RoboDK station: RobotPrint_Printhead_cbeam 1.rdk

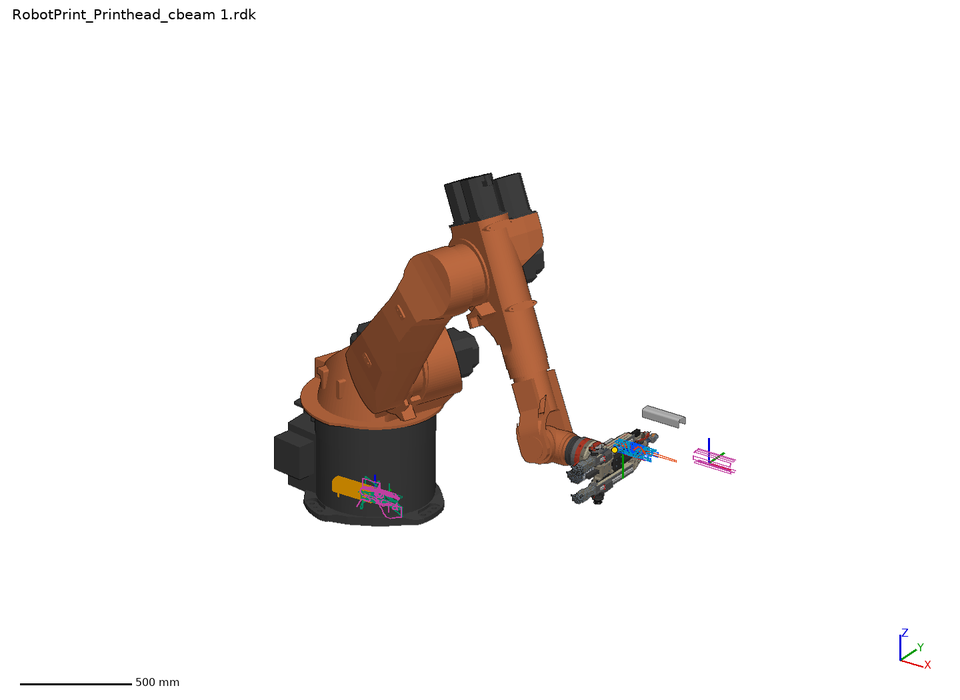
[picture v0: the station drawn from its stored meshes, robots at their saved joint values, targets as dots, program paths as lines]
Station RobotPrinter_Printhead (saved by RoboDK 5.8.0). Poses are relative to the parent item; angles as X-Y-Z fixed-axis rotations.
  - frame KUKA KR 30 HA Base at (0, 0, 0) mm
    - robot KUKA KR 30 HA: 6 axes, payload 30 kg, reach 2033 mm, repeatability 0.05 mm, weight 665 kg
        modified DH rows (alpha deg, a mm, theta deg, d mm): 0, 0, 0, 815; -90, 350, 0, 0; 0, 850, -90, 0; -90, 145, 0, 820; 90, 0, 0, 0; -90, 0, 180, 170
        joint limits [-185, -135, -120, -350, -119, -350] to [185, 35, 158, 350, 119, 350]; home [0, -90, 90, 0, 0, 0]; saved at [20.826, -52.741, 114.474, 203.359, 63.728, -280.823]
      - tool PlasticPos800, TCP at (350.64, -42.92, 173.8) mm
      - tool PlasticPos1200, TCP at (391.44, -42.9, 173.32) mm
      - tool FiberPos800, TCP at (355.38, 32.86, 175) mm, rotated rx 0 ry 90 rz 0 deg
      - tool FiberPos1200, TCP at (394.69, 33.62, 175.94) mm
      - tool Printheady, TCP at (0, 0, 200) mm, size 292.2 x 550.3 x 343.3 mm, geometry from CAD_Printheady.step
      - tool TOOL 0, TCP at (0, 0, 0) mm
    - frame PrintbedOrigin at (1792.66, 35.63, 669.38) mm
    - frame Reference SW at (1415.36, -92.38, 659.99) mm, rotated rx -90 ry 0 rz 0 deg
      - object C-Beam-5mm-200mm RoboDK-Test at (300, -210, 0) mm, size 200 x 40 x 50 mm, geometry from C-Beam-5mm-200mm RoboDK-Test.stl
      - object C-Beam-5mm-200mm RoboDK-Test 1 at (0, 0, 0) mm, size 200 x 50 x 50 mm, geometry from C-Beam-5mm-200mm RoboDK-Test 1.stl
      - object CBL1-2 at (0, 0, 0) mm
      - object CBL2-2 at (0, 0, 0) mm
      - object CBL1 at (0, 0, 0) mm
    - frame BASE 0 at (0, 0, 0) mm
  - machining project CBL1-2 Settings: rotZ(0) | rotX(0)*rotY(0) | onStart | onPathStart | onApproach | onPoint | onRetract | onFinish | SetRPM(%1) | SetTool(%1) | Extruder(%1) | default | default | OutOnMov(%1) | OutOffMov(%1) | onPathFinish | M_RunCode(%1)
  - program CBL1-2 (86 instructions, listed below)
  - machining project CBL2-2 Settings: rotZ(0) | rotX(0)*rotY(0) | rotz(0) | onStart | onPathStart | onApproach | onPoint | onRetract | onFinish | SetRPM(%1) | SetTool(%1) | Extruder(%1) | default | default | OutOnMov(%1) | OutOffMov(%1) | onPathFinish | M_RunCode(%1)
  - program CBL2-2 (24 instructions, listed below)
  - program CBL12 (41 instructions, listed below)
  - program CBL12 (44 instructions, listed below)
  - program CBL12 (39 instructions, listed below)
  - machining project Pfad3 Einstellungen: rotZ(0) | rotX(0)*rotY(0) | onStart | onPathStart | onApproach | onPoint | onRetract | onFinish | SetRPM(%1) | SetTool(%1) | Extruder(%1) | default | default | OutOnMov(%1) | OutOffMov(%1) | onPathFinish | M_RunCode(%1)
  - program Pfad3 (95 instructions, listed below)
  - program TP12Layers (5237 instructions, listed below)
  - machining project CBL1 Settings: rotZ(0) | rotX(0)*rotY(0) | onStart | onPathStart | onApproach | onPoint | onRetract | onFinish | SetRPM(%1) | SetTool(%1) | Extruder(%1) | default | default | OutOnMov(%1) | OutOffMov(%1) | onPathFinish | M_RunCode(%1)
  - program CBL1 (341 instructions, listed below)
  - machining project Pfad5 Einstellungen: rotZ(0) | rotX(0)*rotY(0) | onStart | onPathStart | onApproach | onPoint | onRetract | onFinish | SetRPM(%1) | SetTool(%1) | Extruder(%1) | default | default | OutOnMov(%1) | OutOffMov(%1) | onPathFinish | M_RunCode(%1)
  - program Pfad5 (148 instructions, listed below)
  - machining project Pfad6 Einstellungen: rotZ(0) | rotX(0)*rotY(0) | onStart | onPathStart | onApproach | onPoint | onRetract | onFinish | SetRPM(%1) | SetTool(%1) | Extruder(%1) | default | default | OutOnMov(%1) | OutOffMov(%1) | onPathFinish | M_RunCode(%1)
  - program Pfad6 (33 instructions, listed below)
  - program CFSteer (1006 instructions, listed below)
  - program CFLines (937 instructions, listed below)
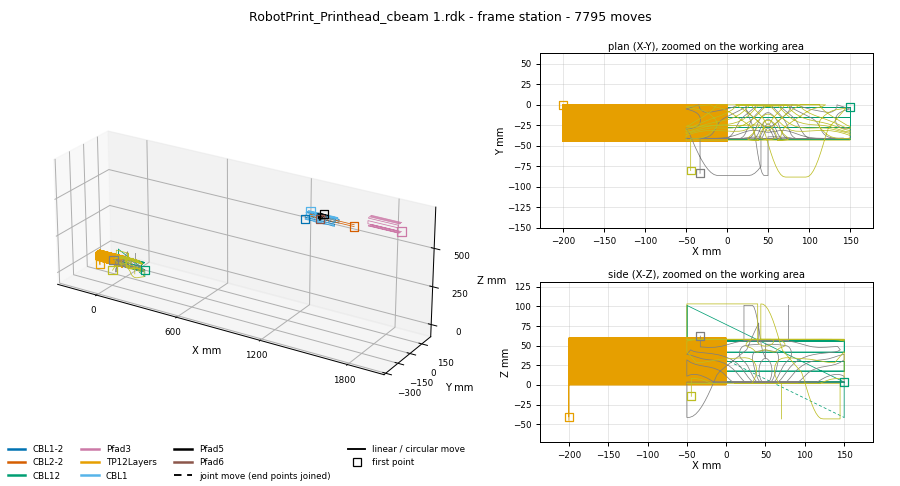
[picture p0: tool path of RobotPrint_Printhead_cbeam 1.rdk in frame station, 7795 of 7795 moves have a stored position in this frame; points joined in program order, loops and branches not executed]

--- program CBL1-2 (robot KUKA KR 30 HA) ---
  Glatt(1)
  Sollgeschwindigkeit (1000.0 mm/s)
  Referenz erstellen.: Reference SW
  Werkzeug setzen: FiberPos800
  Anzeigen FiberPos800
  MoveJ 1 to (-50, -3, 3.75) mm, rotated rx 180 ry 0 rz -90 deg; joints [-10.801, -58.742, 109.357, 0, 39.385, 79.199]
  MoveL 2 to (-50, -3, 3.75) mm, rotated rx 180 ry 0 rz -90 deg; joints [-10.801, -58.742, 109.357, 0, 39.385, 79.199]
  MoveL 3 to (-50, -3, 3.75) mm, rotated rx 180 ry 0 rz -90 deg; joints [-10.801, -58.742, 109.357, 0, 39.385, 79.199]
  MoveL 4 to (-50, -3, 3.75) mm, rotated rx 180 ry 0 rz -90 deg; joints [-10.801, -58.742, 109.357, 0, 39.385, 79.199]
  Sollgeschwindigkeit (50.0 mm/s)
  MoveL 5 to (150, -3, 3.75) mm, rotated rx -180 ry 0 rz -90 deg; joints [-9.475, -48.064, 90.596, 0, 47.468, 80.525]
  Sollgeschwindigkeit (1000.0 mm/s)
  MoveL 6 to (150, -3, 3.75) mm, rotated rx -180 ry 0 rz -90 deg; joints [-9.475, -48.064, 90.596, 0, 47.468, 80.525]
  MoveL 7 to (150, -3, 3.75) mm, rotated rx -180 ry 0 rz -90 deg; joints [-9.475, -48.064, 90.596, 0, 47.468, 80.525]
  Sollgeschwindigkeit (1000.0 mm/s)
  MoveL 8 to (150, -15, 3.75) mm, rotated rx -180 ry 0 rz -90 deg; joints [-9.475, -48.501, 90.408, 0, 48.093, 80.525]
  MoveL 9 to (150, -15, 3.75) mm, rotated rx -180 ry 0 rz -90 deg; joints [-9.475, -48.501, 90.408, 0, 48.093, 80.525]
  MoveL 10 to (150, -15, 3.75) mm, rotated rx -180 ry 0 rz -90 deg; joints [-9.475, -48.501, 90.408, 0, 48.093, 80.525]
  Sollgeschwindigkeit (50.0 mm/s)
  MoveL 11 to (-50, -15, 3.75) mm, rotated rx 180 ry 0 rz -90 deg; joints [-10.801, -59.271, 109.17, 0, 40.102, 79.199]
  Sollgeschwindigkeit (1000.0 mm/s)
  MoveL 12 to (-50, -15, 3.75) mm, rotated rx 180 ry 0 rz -90 deg; joints [-10.801, -59.271, 109.17, 0, 40.102, 79.199]
  MoveL 13 to (-50, -15, 3.75) mm, rotated rx 180 ry 0 rz -90 deg; joints [-10.801, -59.271, 109.17, 0, 40.102, 79.199]
  Sollgeschwindigkeit (1000.0 mm/s)
  MoveL 14 to (-50, -27, 3.75) mm, rotated rx 180 ry 0 rz -90 deg; joints [-10.801, -59.792, 108.97, 0, 40.822, 79.199]
  MoveL 15 to (-50, -27, 3.75) mm, rotated rx 180 ry 0 rz -90 deg; joints [-10.801, -59.792, 108.97, 0, 40.822, 79.199]
  MoveL 16 to (-50, -27, 3.75) mm, rotated rx 180 ry 0 rz -90 deg; joints [-10.801, -59.792, 108.97, 0, 40.822, 79.199]
  Sollgeschwindigkeit (50.0 mm/s)
  MoveL 17 to (150, -27, 3.75) mm, rotated rx -180 ry 0 rz -90 deg; joints [-9.475, -48.931, 90.208, 0, 48.722, 80.525]
  Sollgeschwindigkeit (1000.0 mm/s)
  MoveL 18 to (150, -27, 3.75) mm, rotated rx -180 ry 0 rz -90 deg; joints [-9.475, -48.931, 90.208, 0, 48.722, 80.525]
  MoveL 19 to (150, -27, 3.75) mm, rotated rx -180 ry 0 rz -90 deg; joints [-9.475, -48.931, 90.208, 0, 48.722, 80.525]
  Sollgeschwindigkeit (1000.0 mm/s)
  MoveL 20 to (150, -41.25, 18) mm, rotated rx -180 ry 0 rz -90 deg; joints [-9.972, -49.289, 89.704, 0, 49.585, 80.028]
  MoveL 21 to (150, -41.25, 18) mm, rotated rx -180 ry 0 rz -90 deg; joints [-9.972, -49.289, 89.704, 0, 49.585, 80.028]
  MoveL 22 to (150, -41.25, 18) mm, rotated rx -180 ry 0 rz -90 deg; joints [-9.972, -49.289, 89.704, 0, 49.585, 80.028]
  Sollgeschwindigkeit (50.0 mm/s)
  MoveL 23 to (-50, -41.25, 18) mm, rotated rx -180 ry 0 rz -90 deg; joints [-11.363, -60.254, 108.477, 0, 41.777, 78.637]
  Sollgeschwindigkeit (1000.0 mm/s)
  MoveL 24 to (-50, -41.25, 18) mm, rotated rx -180 ry 0 rz -90 deg; joints [-11.363, -60.254, 108.477, 0, 41.777, 78.637]
  MoveL 25 to (-50, -41.25, 18) mm, rotated rx -180 ry 0 rz -90 deg; joints [-11.363, -60.254, 108.477, 0, 41.777, 78.637]
  Sollgeschwindigkeit (1000.0 mm/s)
  MoveL 26 to (-50, -41.25, 30) mm, rotated rx 180 ry 0 rz -90 deg; joints [-11.835, -60.125, 108.264, 0, 41.86, 78.165]
  MoveL 27 to (-50, -41.25, 30) mm, rotated rx 180 ry 0 rz -90 deg; joints [-11.835, -60.125, 108.264, 0, 41.86, 78.165]
  MoveL 28 to (-50, -41.25, 30) mm, rotated rx 180 ry 0 rz -90 deg; joints [-11.835, -60.125, 108.264, 0, 41.86, 78.165]
  Sollgeschwindigkeit (50.0 mm/s)
  MoveL 29 to (150, -41.25, 30) mm, rotated rx -180 ry 0 rz -90 deg; joints [-10.388, -49.164, 89.482, 0, 49.682, 79.612]
  Sollgeschwindigkeit (1000.0 mm/s)
  MoveL 30 to (150, -41.25, 30) mm, rotated rx -180 ry 0 rz -90 deg; joints [-10.388, -49.164, 89.482, 0, 49.682, 79.612]
  MoveL 31 to (150, -41.25, 30) mm, rotated rx -180 ry 0 rz -90 deg; joints [-10.388, -49.164, 89.482, 0, 49.682, 79.612]
  Sollgeschwindigkeit (1000.0 mm/s)
  MoveL 32 to (150, -41.25, 42) mm, rotated rx 180 ry 0 rz -90 deg; joints [-10.804, -49.033, 89.25, 0, 49.783, 79.196]
  MoveL 33 to (150, -41.25, 42) mm, rotated rx 180 ry 0 rz -90 deg; joints [-10.804, -49.033, 89.25, 0, 49.783, 79.196]
  MoveL 34 to (150, -41.25, 42) mm, rotated rx 180 ry 0 rz -90 deg; joints [-10.804, -49.033, 89.25, 0, 49.783, 79.196]
  Sollgeschwindigkeit (50.0 mm/s)
  MoveL 35 to (-50, -41.25, 42) mm, rotated rx -180 ry 0 rz -90 deg; joints [-12.305, -59.99, 108.043, 0, 41.947, 77.695]
  Sollgeschwindigkeit (1000.0 mm/s)
  MoveL 36 to (-50, -41.25, 42) mm, rotated rx -180 ry 0 rz -90 deg; joints [-12.305, -59.99, 108.043, 0, 41.947, 77.695]
  MoveL 37 to (-50, -41.25, 42) mm, rotated rx -180 ry 0 rz -90 deg; joints [-12.305, -59.99, 108.043, 0, 41.947, 77.695]
  Sollgeschwindigkeit (1000.0 mm/s)
  MoveL 38 to (-50, -27, 56.25) mm, rotated rx 180 ry 0 rz -90 deg; joints [-12.862, -59.222, 108.019, 0, 41.202, 77.138]
  MoveL 39 to (-50, -27, 56.25) mm, rotated rx 180 ry 0 rz -90 deg; joints [-12.862, -59.222, 108.019, 0, 41.202, 77.138]
  MoveL 40 to (-50, -27, 56.25) mm, rotated rx 180 ry 0 rz -90 deg; joints [-12.862, -59.222, 108.019, 0, 41.202, 77.138]
  Sollgeschwindigkeit (50.0 mm/s)
  MoveL 41 to (150, -27, 56.25) mm, rotated rx -180 ry 0 rz -90 deg; joints [-11.296, -48.375, 89.215, 0, 49.16, 78.704]
  Sollgeschwindigkeit (1000.0 mm/s)
  MoveL 42 to (150, -27, 56.25) mm, rotated rx -180 ry 0 rz -90 deg; joints [-11.296, -48.375, 89.215, 0, 49.16, 78.704]
  MoveL 43 to (150, -27, 56.25) mm, rotated rx -180 ry 0 rz -90 deg; joints [-11.296, -48.375, 89.215, 0, 49.16, 78.704]
  Sollgeschwindigkeit (1000.0 mm/s)
  MoveL 44 to (150, -15, 56.25) mm, rotated rx -180 ry 0 rz -90 deg; joints [-11.296, -47.95, 89.416, 0, 48.534, 78.704]
  MoveL 45 to (150, -15, 56.25) mm, rotated rx -180 ry 0 rz -90 deg; joints [-11.296, -47.95, 89.416, 0, 48.534, 78.704]
  MoveL 46 to (150, -15, 56.25) mm, rotated rx -180 ry 0 rz -90 deg; joints [-11.296, -47.95, 89.416, 0, 48.534, 78.704]
  Sollgeschwindigkeit (50.0 mm/s)
  MoveL 47 to (-50, -15, 56.25) mm, rotated rx 180 ry 0 rz -90 deg; joints [-12.862, -58.706, 108.219, 0, 40.488, 77.138]
  Sollgeschwindigkeit (1000.0 mm/s)
  MoveL 48 to (-50, -15, 56.25) mm, rotated rx 180 ry 0 rz -90 deg; joints [-12.862, -58.706, 108.219, 0, 40.488, 77.138]
  MoveL 49 to (-50, -15, 56.25) mm, rotated rx 180 ry 0 rz -90 deg; joints [-12.862, -58.706, 108.219, 0, 40.488, 77.138]
  Sollgeschwindigkeit (1000.0 mm/s)
  MoveL 50 to (-50, -3, 56.25) mm, rotated rx 180 ry 0 rz -90 deg; joints [-12.862, -58.183, 108.406, 0, 39.777, 77.138]
  MoveL 51 to (-50, -3, 56.25) mm, rotated rx 180 ry 0 rz -90 deg; joints [-12.862, -58.183, 108.406, 0, 39.777, 77.138]
  MoveL 52 to (-50, -3, 56.25) mm, rotated rx 180 ry 0 rz -90 deg; joints [-12.862, -58.183, 108.406, 0, 39.777, 77.138]
  Sollgeschwindigkeit (50.0 mm/s)
  MoveL 53 to (150, -3, 56.25) mm, rotated rx -180 ry 0 rz -90 deg; joints [-11.296, -47.517, 89.605, 0, 47.912, 78.704]
  Sollgeschwindigkeit (1000.0 mm/s)
  MoveL 54 to (150, -3, 56.25) mm, rotated rx -180 ry 0 rz -90 deg; joints [-11.296, -47.517, 89.605, 0, 47.912, 78.704]
  MoveL 55 to (150, -3, 56.25) mm, rotated rx -180 ry 0 rz -90 deg; joints [-11.296, -47.517, 89.605, 0, 47.912, 78.704]

--- program CBL2-2 (robot KUKA KR 30 HA) ---
  Glatt(1)
  Sollgeschwindigkeit (1000.0 mm/s)
  Referenz erstellen.: Reference SW
  Werkzeug setzen: FiberPos800
  Anzeigen FiberPos800
  MoveJ 1 to (250, -3, 58.75) mm, rotated rx 90 ry 0 rz -90 deg; joints [1.885, -7.943, 13.331, 0, 84.613, 1.885]
  MoveL 2 to (250, -3, 58.75) mm, rotated rx 90 ry 0 rz -90 deg; joints [1.885, -7.943, 13.331, 0, 84.613, 1.885]
  MoveL 3 to (150, -3, 58.75) mm, rotated rx 90 ry 0 rz -90 deg; joints [1.983, -26.347, 49.734, 0, 66.613, 1.983]
  MoveL 4 to (150, -3, 58.75) mm, rotated rx 90 ry 0 rz -90 deg; joints [1.983, -26.347, 49.734, 0, 66.613, 1.983]
  Sollgeschwindigkeit (50.0 mm/s)
  MoveL 5 to (-50, -3, 58.75) mm, rotated rx 90 ry 0 rz -90 deg; joints [2.213, -41.91, 79.315, 0, 52.595, 2.213]
  Sollgeschwindigkeit (1000.0 mm/s)
  MoveL 6 to (-50, -3, 58.75) mm, rotated rx 90 ry 0 rz -90 deg; joints [2.213, -41.91, 79.315, 0, 52.595, 2.213]
  MoveL 7 to (50, -3, 58.75) mm, rotated rx 90 ry 0 rz -90 deg; joints [2.091, -35.006, 66.355, 0, 58.651, 2.091]
  Sollgeschwindigkeit (1000.0 mm/s)
  MoveL 8 to (50, -15, 58.75) mm, rotated rx 90 ry 0 rz -90 deg; joints [2.091, -35.355, 66.132, 0, 59.223, 2.091]
  MoveL 9 to (-50, -15, 58.75) mm, rotated rx 90 ry 0 rz -90 deg; joints [2.213, -42.303, 79.116, 0, 53.187, 2.213]
  MoveL 10 to (-50, -15, 58.75) mm, rotated rx 90 ry 0 rz -90 deg; joints [2.213, -42.303, 79.116, 0, 53.187, 2.213]
  Sollgeschwindigkeit (50.0 mm/s)
  MoveL 11 to (150, -15, 58.75) mm, rotated rx 90 ry 0 rz -90 deg; joints [1.983, -26.634, 49.443, 0, 67.192, 1.983]
  Sollgeschwindigkeit (1000.0 mm/s)
  MoveL 12 to (150, -15, 58.75) mm, rotated rx 90 ry 0 rz -90 deg; joints [1.983, -26.634, 49.443, 0, 67.192, 1.983]
  MoveL 13 to (250, -15, 58.75) mm, rotated rx 90 ry -20 rz -90 deg; joints [-1.516, -8.156, 13.591, 20.06, 85.412, -3.287]
  Sollgeschwindigkeit (1000.0 mm/s)

--- program CBL12 (robot KUKA KR 30 HA) ---
  BAS (#INITMOV,0)
  BAS (#VEL_PTP,100)
  BAS (#ACC_PTP,20)
  Sollgeschwindigkeit (200.0 mm/s)
  Werkzeug setzen: TOOL 0
  Referenz erstellen.: BASE 0
  $ADVANCE = 5
  $APO.CPTP = 1.000
  $APO.CDIS = 1.000
  Sollgeschwindigkeit (1000.0 mm/s)
  Frame wechseln at (1415.36, -92.38, 651.84) mm, rotated rx -90 ry 0 rz 0 deg
  Werkzeug setzen at (355.38, 32.86, 175) mm, rotated rx 0 ry 90 rz 0 deg
  Sollgeschwindigkeit (50.0 mm/s)
  Sollgeschwindigkeit (50.0 mm/s)
  MoveL 2 to (150, -3, 3.75) mm, rotated rx 0 ry 0 rz 180 deg; joints [19.993, -42.546, 119.796, -159.543, 78.03, 85.576]
  MoveL 3 to (-50, -3, 3.75) mm, rotated rx 0 ry 0 rz 180 deg; joints [23.516, -46.815, 134.283, -156.463, 87.679, 88.989]
  MoveL 4 to (-50, -15, 3.75) mm, rotated rx 0 ry 0 rz 180 deg; joints [23.516, -47.77, 134.503, -156.449, 87.005, 88.695]
  MoveL 5 to (150, -15, 3.75) mm, rotated rx 0 ry 0 rz 180 deg; joints [19.993, -43.337, 119.989, -159.497, 77.47, 85.362]
  MoveL 6 to (150, -27, 3.75) mm, rotated rx 0 ry 0 rz 180 deg; joints [19.993, -44.126, 120.17, -159.449, 76.901, 85.143]
  MoveL 7 to (-50, -27, 3.75) mm, rotated rx 0 ry 0 rz 180 deg; joints [23.516, -48.725, 134.71, -156.432, 86.319, 88.396]
  MoveL 8 to (-50, -30, 3.75) mm, rotated rx 0 ry 0 rz 180 deg; joints [23.516, -48.963, 134.759, -156.427, 86.146, 88.32]
  MoveL 9 to (-50, -35.62, 5.26) mm, rotated rx 30 ry 0 rz 180 deg; joints [21.955, -63.996, 137.068, -157.151, 74.333, 113.508]
  MoveL 10 to (-50, -39.74, 9.38) mm, rotated rx 60 ry 0 rz 180 deg; joints [15.822, -76.367, 138.611, -162.243, 63.381, 141.835]
  MoveL 11 to (-50, -41.25, 15) mm, rotated rx 90 ry 0 rz 180 deg; joints [6.167, -82.637, 139.716, -172.666, 57.294, 176.022]
  MoveL 12 to (-50, -41.25, 18) mm, rotated rx 90 ry 0 rz 180 deg; joints [6, -82.656, 139.739, -172.863, 57.286, 176.129]
  MoveL 13 to (150, -41.25, 18) mm, rotated rx 90 ry 0 rz 180 deg; joints [5.022, -71.46, 124.912, -173.757, 53.616, 176.287]
  MoveL 14 to (150, -41.25, 30) mm, rotated rx 90 ry 0 rz 180 deg; joints [4.463, -71.513, 124.99, -174.453, 53.605, 176.702]
  MoveL 15 to (-50, -41.25, 30) mm, rotated rx 90 ry 0 rz 180 deg; joints [5.333, -82.727, 139.823, -173.656, 57.257, 176.559]
  MoveL 16 to (-50, -41.25, 42) mm, rotated rx 90 ry 0 rz 180 deg; joints [4.664, -82.789, 139.898, -174.451, 57.231, 176.99]
  MoveL 17 to (150, -41.25, 42) mm, rotated rx 90 ry 0 rz 180 deg; joints [3.902, -71.56, 125.058, -175.15, 53.596, 177.117]
  MoveL 18 to (150, -41.25, 45) mm, rotated rx 90 ry 0 rz 180 deg; joints [3.762, -71.571, 125.074, -175.324, 53.594, 177.221]
  MoveL 19 to (150, -39.74, 50.62) mm, rotated rx 120 ry 0 rz 180 deg; joints [-5.033, -69.749, 125.546, 173.922, 55.947, -146.588]
  MoveL 20 to (150, -35.62, 54.74) mm, rotated rx 150 ry 0 rz 180 deg; joints [-11.744, -61.757, 125.379, 166.936, 64.215, -114.236]
  MoveL 21 to (150, -30, 56.25) mm, rotated rx 180 ry 0 rz 180 deg; joints [-14.66, -49.801, 124, 164.79, 74.727, -85.904]
  MoveL 22 to (150, -27, 56.25) mm, rotated rx 180 ry 0 rz 180 deg; joints [-14.66, -49.601, 123.973, 164.803, 74.893, -85.95]
  MoveL 23 to (-50, -27, 56.25) mm, rotated rx 180 ry 0 rz 180 deg; joints [-17.374, -55.024, 138.883, 162.532, 84.14, -88.16]
  MoveL 24 to (-50, -15, 56.25) mm, rotated rx 180 ry 0 rz 180 deg; joints [-17.374, -54.025, 138.747, 162.557, 84.963, -88.42]
  MoveL 25 to (150, -15, 56.25) mm, rotated rx 180 ry 0 rz 180 deg; joints [-14.66, -48.802, 123.857, 164.85, 75.553, -86.135]
  MoveL 26 to (150, -3, 56.25) mm, rotated rx 180 ry 0 rz 180 deg; joints [-14.66, -47.998, 123.728, 164.894, 76.204, -86.317]
  MoveL 27 to (-50, -3, 56.25) mm, rotated rx 180 ry 0 rz 180 deg; joints [-17.374, -53.024, 138.596, 162.577, 85.774, -88.675]
  END

--- program CBL12 (robot KUKA KR 30 HA) ---
  BAS (#INITMOV,0)
  BAS (#VEL_PTP,100)
  BAS (#ACC_PTP,20)
  Sollgeschwindigkeit (200.0 mm/s)
  Werkzeug setzen: TOOL 0
  Referenz erstellen.: BASE 0
  $ADVANCE = 5
  $APO.CPTP = 1.000
  $APO.CDIS = 1.000
  Sollgeschwindigkeit (1000.0 mm/s)
  Frame wechseln at (1415.36, -92.38, 651.84) mm, rotated rx -90 ry 0 rz 0 deg
  Werkzeug setzen at (355.38, 32.86, 175) mm, rotated rx 0 ry 90 rz 0 deg
  MoveJ 1 to (150, -3, -41.25) mm, rotated rx 0 ry 0 rz 180 deg; joints [21.837, -42.094, 118.479, -157.594, 77.378, 84.852]
  Sollgeschwindigkeit (50.0 mm/s)
  MoveL 2 to (150, -3, 3.75) mm, rotated rx 0 ry 0 rz 180 deg; joints [19.993, -42.546, 119.796, -159.543, 78.03, 85.576]
  Sollgeschwindigkeit (50.0 mm/s)
  MoveL 3 to (-50, -3, 3.75) mm, rotated rx 0 ry 0 rz 180 deg; joints [23.516, -46.815, 134.283, -156.463, 87.679, 88.989]
  MoveL 4 to (-50, -15, 3.75) mm, rotated rx 0 ry 0 rz 180 deg; joints [23.516, -47.77, 134.503, -156.449, 87.005, 88.695]
  MoveL 5 to (150, -15, 3.75) mm, rotated rx 0 ry 0 rz 180 deg; joints [19.993, -43.337, 119.989, -159.497, 77.47, 85.362]
  MoveL 6 to (150, -27, 3.75) mm, rotated rx 0 ry 0 rz 180 deg; joints [19.993, -44.126, 120.17, -159.449, 76.901, 85.143]
  MoveL 7 to (-50, -27, 3.75) mm, rotated rx 0 ry 0 rz 180 deg; joints [23.516, -48.725, 134.71, -156.432, 86.319, 88.396]
  MoveL 8 to (-50, -30, 3.75) mm, rotated rx 0 ry 0 rz 180 deg; joints [23.516, -48.963, 134.759, -156.427, 86.146, 88.32]
  MoveL 9 to (-50, -35.62, 5.26) mm, rotated rx 30 ry 0 rz 180 deg; joints [21.955, -63.996, 137.068, -157.151, 74.333, 113.508]
  MoveL 10 to (-50, -39.74, 9.38) mm, rotated rx 60 ry 0 rz 180 deg; joints [15.822, -76.367, 138.611, -162.243, 63.381, 141.835]
  MoveL 11 to (-50, -41.25, 15) mm, rotated rx 90 ry 0 rz 180 deg; joints [6.167, -82.637, 139.716, -172.666, 57.294, 176.022]
  MoveL 12 to (-50, -41.25, 18) mm, rotated rx 90 ry 0 rz 180 deg; joints [6, -82.656, 139.739, -172.863, 57.286, 176.129]
  MoveL 13 to (150, -41.25, 18) mm, rotated rx 90 ry 0 rz 180 deg; joints [5.022, -71.46, 124.912, -173.757, 53.616, 176.287]
  MoveL 14 to (150, -41.25, 30) mm, rotated rx 90 ry 0 rz 180 deg; joints [4.463, -71.513, 124.99, -174.453, 53.605, 176.702]
  MoveL 15 to (-50, -41.25, 30) mm, rotated rx 90 ry 0 rz 180 deg; joints [5.333, -82.727, 139.823, -173.656, 57.257, 176.559]
  MoveL 16 to (-50, -41.25, 42) mm, rotated rx 90 ry 0 rz 180 deg; joints [4.664, -82.789, 139.898, -174.451, 57.231, 176.99]
  MoveL 17 to (150, -41.25, 42) mm, rotated rx 90 ry 0 rz 180 deg; joints [3.902, -71.56, 125.058, -175.15, 53.596, 177.117]
  MoveL 18 to (150, -41.25, 45) mm, rotated rx 90 ry 0 rz 180 deg; joints [3.762, -71.571, 125.074, -175.324, 53.594, 177.221]
  MoveL 19 to (150, -39.74, 50.62) mm, rotated rx 120 ry 0 rz 180 deg; joints [-5.033, -69.749, 125.546, 173.922, 55.947, -146.588]
  MoveL 20 to (150, -35.62, 54.74) mm, rotated rx 150 ry 0 rz 180 deg; joints [-11.744, -61.757, 125.379, 166.936, 64.215, -114.236]
  MoveL 21 to (150, -30, 56.25) mm, rotated rx 180 ry 0 rz 180 deg; joints [-14.66, -49.801, 124, 164.79, 74.727, -85.904]
  MoveL 22 to (150, -27, 56.25) mm, rotated rx 180 ry 0 rz 180 deg; joints [-14.66, -49.601, 123.973, 164.803, 74.893, -85.95]
  MoveL 23 to (-50, -27, 56.25) mm, rotated rx 180 ry 0 rz 180 deg; joints [-17.374, -55.024, 138.883, 162.532, 84.14, -88.16]
  MoveL 24 to (-50, -15, 56.25) mm, rotated rx 180 ry 0 rz 180 deg; joints [-17.374, -54.025, 138.747, 162.557, 84.963, -88.42]
  MoveL 25 to (150, -15, 56.25) mm, rotated rx 180 ry 0 rz 180 deg; joints [-14.66, -48.802, 123.857, 164.85, 75.553, -86.135]
  MoveL 26 to (150, -3, 56.25) mm, rotated rx 180 ry 0 rz 180 deg; joints [-14.66, -47.998, 123.728, 164.894, 76.204, -86.317]
  MoveL 27 to (-50, -3, 56.25) mm, rotated rx 180 ry 0 rz 180 deg; joints [-17.374, -53.024, 138.596, 162.577, 85.774, -88.675]
  Sollgeschwindigkeit (1000.0 mm/s)
  MoveL 28 to (-50, -3, 101.25) mm, rotated rx 180 ry 0 rz 180 deg; joints [-19.645, -52.711, 137.529, 160.28, 85.121, -88.254]
  END

--- program CBL12 (robot KUKA KR 30 HA) ---
  BAS (#INITMOV,0)
  BAS (#VEL_PTP,100)
  BAS (#ACC_PTP,20)
  Sollgeschwindigkeit (200.0 mm/s)
  Werkzeug setzen: TOOL 0
  Referenz erstellen.: BASE 0
  $ADVANCE = 5
  $APO.CPTP = 1.000
  $APO.CDIS = 1.000
  Sollgeschwindigkeit (1000.0 mm/s)
  Frame wechseln at (1415.36, -92.38, 651.84) mm, rotated rx -90 ry 0 rz 0 deg
  Werkzeug setzen at (355.38, 32.86, 175) mm, rotated rx 0 ry 90 rz 0 deg
  Sollgeschwindigkeit (50.0 mm/s)
  MoveL 2 to (150, -3, 3.75) mm, rotated rx 0 ry 0 rz 180 deg; joints [19.993, -42.546, 119.796, -159.543, 78.03, 85.576]
  Sollgeschwindigkeit (50.0 mm/s)
  MoveL 3 to (-50, -3, 3.75) mm, rotated rx 0 ry 0 rz 180 deg; joints [23.516, -46.815, 134.283, -156.463, 87.679, 88.989]
  MoveL 4 to (-50, -15, 3.75) mm, rotated rx 0 ry 0 rz 180 deg; joints [23.516, -47.77, 134.503, -156.449, 87.005, 88.695]
  MoveL 5 to (150, -15, 3.75) mm, rotated rx 0 ry 0 rz 180 deg; joints [19.993, -43.337, 119.989, -159.497, 77.47, 85.362]
  MoveL 6 to (150, -27, 3.75) mm, rotated rx 0 ry 0 rz 180 deg; joints [19.993, -44.126, 120.17, -159.449, 76.901, 85.143]
  MoveL 7 to (-50, -27, 3.75) mm, rotated rx 0 ry 0 rz 180 deg; joints [23.516, -48.725, 134.71, -156.432, 86.319, 88.396]
  MoveL 8 to (-50, -30, 3.75) mm, rotated rx 0 ry 0 rz 180 deg; joints [23.516, -48.963, 134.759, -156.427, 86.146, 88.32]
  MoveC to (-50, -37.95, 6.71) mm, rotated rx 45 ry 0 rz 180 deg; joints [19.444, -70.739, 137.919, -159.043, 68.547, 127.026] to (-50, -41.25, 15) mm, rotated rx 90 ry 0 rz 180 deg; joints [6.167, -82.637, 139.716, -172.666, 57.294, 176.022]
  MoveL 10 to (-50, -41.25, 18) mm, rotated rx 90 ry 0 rz 180 deg; joints [6, -82.656, 139.739, -172.863, 57.286, 176.129]
  MoveL 11 to (150, -41.25, 18) mm, rotated rx 90 ry 0 rz 180 deg; joints [5.022, -71.46, 124.912, -173.757, 53.616, 176.287]
  MoveL 12 to (150, -41.25, 30) mm, rotated rx 90 ry 0 rz 180 deg; joints [4.463, -71.513, 124.99, -174.453, 53.605, 176.702]
  MoveL 13 to (-50, -41.25, 30) mm, rotated rx 90 ry 0 rz 180 deg; joints [5.333, -82.727, 139.823, -173.656, 57.257, 176.559]
  MoveL 14 to (-50, -41.25, 42) mm, rotated rx 90 ry 0 rz 180 deg; joints [4.664, -82.789, 139.898, -174.451, 57.231, 176.99]
  MoveL 15 to (150, -41.25, 42) mm, rotated rx 90 ry 0 rz 180 deg; joints [3.902, -71.56, 125.058, -175.15, 53.596, 177.117]
  MoveL 16 to (150, -41.25, 45) mm, rotated rx 90 ry 0 rz 180 deg; joints [3.762, -71.571, 125.074, -175.324, 53.594, 177.221]
  MoveC to (150, -37.95, 53.3) mm, rotated rx 135 ry 0 rz 180 deg; joints [-8.802, -66.42, 125.579, -190.223, 59.561, 230.221] to (150, -30, 56.25) mm, rotated rx 180 ry 0 rz 180 deg; joints [-14.66, -49.801, 124, -195.21, 74.727, 274.096]
  MoveL 18 to (150, -27, 56.25) mm, rotated rx 180 ry 0 rz 180 deg; joints [-14.66, -49.601, 123.973, 164.803, 74.893, -85.95]
  MoveL 19 to (-50, -27, 56.25) mm, rotated rx 180 ry 0 rz 180 deg; joints [-17.374, -55.024, 138.883, 162.532, 84.14, -88.16]
  MoveL 20 to (-50, -15, 56.25) mm, rotated rx 180 ry 0 rz 180 deg; joints [-17.374, -54.025, 138.747, 162.557, 84.963, -88.42]
  MoveL 21 to (150, -15, 56.25) mm, rotated rx 180 ry 0 rz 180 deg; joints [-14.66, -48.802, 123.857, 164.85, 75.553, -86.135]
  MoveL 22 to (150, -3, 56.25) mm, rotated rx 180 ry 0 rz 180 deg; joints [-14.66, -47.998, 123.728, 164.894, 76.204, -86.317]
  MoveL 23 to (-50, -3, 56.25) mm, rotated rx 180 ry 0 rz 180 deg; joints [-17.374, -53.024, 138.596, 162.577, 85.774, -88.675]
  Sollgeschwindigkeit (50.0 mm/s)
  MoveL 24 to (-50, -3, 101.25) mm, rotated rx 180 ry 0 rz 180 deg; joints [-19.645, -52.711, 137.529, 160.28, 85.121, -88.254]
  END

--- program Pfad3 (robot KUKA KR 30 HA) ---
  Glatt(1)
  Sollgeschwindigkeit (1000.0 mm/s)
  Referenz erstellen.: PrintbedOrigin
  Werkzeug setzen: PlasticPos800
  Anzeigen PlasticPos800
  MoveJ 1 to (150, -3, 1.25) mm; joints [19.7, -42.107, 120.306, -70.685, 93.953, -101.127]
  MoveL 2 to (150, -3, 1.25) mm; joints [19.7, -42.107, 120.306, -70.685, 93.953, -101.127]
  MoveL 3 to (150, -3, 1.25) mm; joints [19.7, -42.107, 120.306, -70.685, 93.953, -101.127]
  MoveL 4 to (150, -3, 1.25) mm; joints [19.7, -42.107, 120.306, -70.685, 93.953, -101.127]
  Sollgeschwindigkeit (50.0 mm/s)
  MoveL 5 to (-50, -3, 1.25) mm; joints [23.201, -46.159, 134.741, -66.805, 90.559, -91.303]
  Sollgeschwindigkeit (1000.0 mm/s)
  MoveL 6 to (-50, -3, 1.25) mm; joints [23.201, -46.159, 134.741, -66.805, 90.559, -91.303]
  MoveL 7 to (-50, -3, 1.25) mm; joints [23.201, -46.159, 134.741, -66.805, 90.559, -91.303]
  Sollgeschwindigkeit (1000.0 mm/s)
  MoveL 8 to (-50, -15, 1.25) mm; joints [23.201, -47.124, 134.975, -66.814, 90.847, -91.976]
  MoveL 9 to (-50, -15, 1.25) mm; joints [23.201, -47.124, 134.975, -66.814, 90.847, -91.976]
  MoveL 10 to (-50, -15, 1.25) mm; joints [23.201, -47.124, 134.975, -66.814, 90.847, -91.976]
  Sollgeschwindigkeit (50.0 mm/s)
  MoveL 11 to (150, -15, 1.25) mm; joints [19.7, -42.906, 120.511, -70.725, 94.15, -101.69]
  Sollgeschwindigkeit (1000.0 mm/s)
  MoveL 12 to (150, -15, 1.25) mm; joints [19.7, -42.906, 120.511, -70.725, 94.15, -101.69]
  MoveL 13 to (150, -15, 1.25) mm; joints [19.7, -42.906, 120.511, -70.725, 94.15, -101.69]
  Sollgeschwindigkeit (1000.0 mm/s)
  MoveL 14 to (150, -27, 1.25) mm; joints [19.7, -43.703, 120.703, -70.767, 94.349, -102.263]
  MoveL 15 to (150, -27, 1.25) mm; joints [19.7, -43.703, 120.703, -70.767, 94.349, -102.263]
  MoveL 16 to (150, -27, 1.25) mm; joints [19.7, -43.703, 120.703, -70.767, 94.349, -102.263]
  Sollgeschwindigkeit (50.0 mm/s)
  MoveL 17 to (-50, -27, 1.25) mm; joints [23.201, -48.089, 135.194, -66.825, 91.14, -92.661]
  Sollgeschwindigkeit (1000.0 mm/s)
  MoveL 18 to (-50, -27, 1.25) mm; joints [23.201, -48.089, 135.194, -66.825, 91.14, -92.661]
  MoveL 19 to (-50, -27, 1.25) mm; joints [23.201, -48.089, 135.194, -66.825, 91.14, -92.661]
  Sollgeschwindigkeit (1000.0 mm/s)
  MoveL 20 to (-50, -39.72, 5.28) mm; joints [23.009, -49.142, 135.53, -67.032, 91.411, -93.325]
  MoveL 21 to (-50, -39.72, 5.28) mm; joints [23.009, -49.142, 135.53, -67.032, 91.411, -93.325]
  MoveL 22 to (-50, -39.72, 5.28) mm; joints [23.009, -49.142, 135.53, -67.032, 91.411, -93.325]
  Sollgeschwindigkeit (50.0 mm/s)
  MoveL 23 to (150, -39.72, 5.28) mm; joints [19.531, -44.584, 121.003, -70.975, 94.503, -102.826]
  Sollgeschwindigkeit (1000.0 mm/s)
  MoveL 24 to (150, -39.72, 5.28) mm; joints [19.531, -44.584, 121.003, -70.975, 94.503, -102.826]
  MoveL 25 to (150, -39.72, 5.28) mm; joints [19.531, -44.584, 121.003, -70.975, 94.503, -102.826]
  Sollgeschwindigkeit (1000.0 mm/s)
  MoveL 26 to (150, -43.75, 20) mm; joints [18.912, -44.991, 121.455, -71.577, 94.351, -102.831]
  MoveL 27 to (150, -43.75, 20) mm; joints [18.912, -44.991, 121.455, -71.577, 94.351, -102.831]
  MoveL 28 to (150, -43.75, 20) mm; joints [18.912, -44.991, 121.455, -71.577, 94.351, -102.831]
  Sollgeschwindigkeit (50.0 mm/s)
  MoveL 29 to (-50, -43.75, 20) mm; joints [22.301, -49.578, 136.02, -67.738, 91.349, -93.292]
  Sollgeschwindigkeit (1000.0 mm/s)
  MoveL 30 to (-50, -43.75, 20) mm; joints [22.301, -49.578, 136.02, -67.738, 91.349, -93.292]
  MoveL 31 to (-50, -43.75, 20) mm; joints [22.301, -49.578, 136.02, -67.738, 91.349, -93.292]
  Sollgeschwindigkeit (1000.0 mm/s)
  MoveL 32 to (-50, -43.75, 40) mm; joints [21.327, -49.721, 136.575, -68.702, 91.144, -92.932]
  MoveL 33 to (-50, -43.75, 40) mm; joints [21.327, -49.721, 136.575, -68.702, 91.144, -92.932]
  MoveL 34 to (-50, -43.75, 40) mm; joints [21.327, -49.721, 136.575, -68.702, 91.144, -92.932]
  Sollgeschwindigkeit (50.0 mm/s)
  MoveL 35 to (150, -43.75, 40) mm; joints [18.064, -45.174, 121.969, -72.384, 94.062, -102.575]
  Sollgeschwindigkeit (1000.0 mm/s)
  MoveL 36 to (150, -43.75, 40) mm; joints [18.064, -45.174, 121.969, -72.384, 94.062, -102.575]
  MoveL 37 to (150, -43.75, 40) mm; joints [18.064, -45.174, 121.969, -72.384, 94.062, -102.575]
  Sollgeschwindigkeit (1000.0 mm/s)
  MoveL 38 to (150, -39.72, 54.72) mm; joints [17.434, -45.032, 122.274, -72.971, 93.794, -102.19]
  MoveL 39 to (150, -39.72, 54.72) mm; joints [17.434, -45.032, 122.274, -72.971, 93.794, -102.19]
  MoveL 40 to (150, -39.72, 54.72) mm; joints [17.434, -45.032, 122.274, -72.971, 93.794, -102.19]
  Sollgeschwindigkeit (50.0 mm/s)
  MoveL 41 to (-50, -39.72, 54.72) mm; joints [20.603, -49.49, 136.9, -69.417, 90.911, -92.425]
  Sollgeschwindigkeit (1000.0 mm/s)
  MoveL 42 to (-50, -39.72, 54.72) mm; joints [20.603, -49.49, 136.9, -69.417, 90.911, -92.425]
  MoveL 43 to (-50, -39.72, 54.72) mm; joints [20.603, -49.49, 136.9, -69.417, 90.911, -92.425]
  Sollgeschwindigkeit (1000.0 mm/s)
  MoveL 44 to (-50, -27, 58.75) mm; joints [20.403, -48.468, 136.782, -69.605, 90.588, -91.58]
  MoveL 45 to (-50, -27, 58.75) mm; joints [20.403, -48.468, 136.782, -69.605, 90.588, -91.58]
  MoveL 46 to (-50, -27, 58.75) mm; joints [20.403, -48.468, 136.782, -69.605, 90.588, -91.58]
  Sollgeschwindigkeit (50.0 mm/s)
  MoveL 47 to (150, -27, 58.75) mm; joints [17.261, -44.209, 122.179, -73.096, 93.546, -101.503]
  Sollgeschwindigkeit (1000.0 mm/s)
  MoveL 48 to (150, -27, 58.75) mm; joints [17.261, -44.209, 122.179, -73.096, 93.546, -101.503]
  MoveL 49 to (150, -27, 58.75) mm; joints [17.261, -44.209, 122.179, -73.096, 93.546, -101.503]
  Sollgeschwindigkeit (1000.0 mm/s)
  MoveL 50 to (150, -15, 58.75) mm; joints [17.261, -43.398, 121.985, -73.061, 93.366, -100.912]
  MoveL 51 to (150, -15, 58.75) mm; joints [17.261, -43.398, 121.985, -73.061, 93.366, -100.912]
  MoveL 52 to (150, -15, 58.75) mm; joints [17.261, -43.398, 121.985, -73.061, 93.366, -100.912]
  Sollgeschwindigkeit (50.0 mm/s)
  MoveL 53 to (-50, -15, 58.75) mm; joints [20.403, -47.48, 136.558, -69.599, 90.321, -90.864]
  Sollgeschwindigkeit (1000.0 mm/s)
  MoveL 54 to (-50, -15, 58.75) mm; joints [20.403, -47.48, 136.558, -69.599, 90.321, -90.864]
  MoveL 55 to (-50, -15, 58.75) mm; joints [20.403, -47.48, 136.558, -69.599, 90.321, -90.864]
  Sollgeschwindigkeit (1000.0 mm/s)
  MoveL 56 to (-50, -3, 58.75) mm; joints [20.403, -46.492, 136.32, -69.597, 90.06, -90.161]
  MoveL 57 to (-50, -3, 58.75) mm; joints [20.403, -46.492, 136.32, -69.597, 90.06, -90.161]
  MoveL 58 to (-50, -3, 58.75) mm; joints [20.403, -46.492, 136.32, -69.597, 90.06, -90.161]
  Sollgeschwindigkeit (50.0 mm/s)
  MoveL 59 to (150, -3, 58.75) mm; joints [17.261, -42.586, 121.778, -73.028, 93.189, -100.331]
  Sollgeschwindigkeit (1000.0 mm/s)
  MoveL 60 to (150, -3, 58.75) mm; joints [17.261, -42.586, 121.778, -73.028, 93.189, -100.331]
  MoveL 61 to (150, -3, 58.75) mm; joints [17.261, -42.586, 121.778, -73.028, 93.189, -100.331]

--- program TP12Layers (robot KUKA KR 30 HA) ---
  BAS (#INITMOV,0)
  BAS (#VEL_PTP,100)
  BAS (#ACC_PTP,20)
  Sollgeschwindigkeit (200.0 mm/s)
  Werkzeug setzen: TOOL 0
  Referenz erstellen.: BASE 0
  $ADVANCE = 5
  $APO.CPTP = 1.000
  $APO.CDIS = 1.000
  Sollgeschwindigkeit (1000.0 mm/s)
  Frame wechseln at (1715.36, -93.32, 871.24) mm, rotated rx -90 ry 0 rz 0 deg
  Werkzeug setzen at (357.66, -43.21, 173.4) mm, rotated rx 0 ry 90 rz 0 deg
  MoveJ 2 to (-200, 0, -40.4) mm, rotated rx 0 ry 0 rz 180 deg; joints [22.747, -61.882, 123.249, -154.466, 63.773, 78.079]
  Sollgeschwindigkeit (25.0 mm/s)
  MoveL 3 to (-200, 0, 4.6) mm, rotated rx 0 ry 0 rz 180 deg; joints [20.851, -62.647, 124.599, -156.656, 63.933, 79.262]
  MoveL 4 to (0, 0, 4.6) mm, rotated rx 0 ry 0 rz 180 deg; joints [18.023, -53.821, 108.638, -158.293, 56.776, 77.695]
  MoveL 5 to (0, -0.6, 4.6) mm, rotated rx 0 ry 0 rz 180 deg; joints [18.023, -53.85, 108.633, -158.285, 56.744, 77.681]
  MoveL 6 to (-200, -0.6, 4.6) mm, rotated rx 0 ry 0 rz 180 deg; joints [20.851, -62.682, 124.594, -156.649, 63.896, 79.244]
  MoveL 7 to (-200, -1.2, 4.6) mm, rotated rx 0 ry 0 rz 180 deg; joints [20.851, -62.717, 124.588, -156.641, 63.859, 79.226]
  MoveL 8 to (0, -1.2, 4.6) mm, rotated rx 0 ry 0 rz 180 deg; joints [18.023, -53.879, 108.628, -158.277, 56.713, 77.666]
  MoveL 9 to (0, -1.8, 4.6) mm, rotated rx 0 ry 0 rz 180 deg; joints [18.023, -53.907, 108.623, -158.269, 56.682, 77.651]
  MoveL 10 to (-200, -1.8, 4.6) mm, rotated rx 0 ry 0 rz 180 deg; joints [20.851, -62.752, 124.583, -156.633, 63.822, 79.209]
  MoveL 11 to (-200, -2.4, 4.6) mm, rotated rx 0 ry 0 rz 180 deg; joints [20.851, -62.787, 124.578, -156.625, 63.785, 79.191]
  MoveL 12 to (0, -2.4, 4.6) mm, rotated rx 0 ry 0 rz 180 deg; joints [18.023, -53.936, 108.618, -158.26, 56.65, 77.636]
  MoveL 13 to (0, -3, 4.6) mm, rotated rx 0 ry 0 rz 180 deg; joints [18.023, -53.965, 108.613, -158.252, 56.619, 77.621]
  MoveL 14 to (-200, -3, 4.6) mm, rotated rx 0 ry 0 rz 180 deg; joints [20.851, -62.822, 124.572, -156.617, 63.748, 79.173]
  MoveL 15 to (-200, -3.6, 4.6) mm, rotated rx 0 ry 0 rz 180 deg; joints [20.851, -62.857, 124.567, -156.609, 63.711, 79.155]
  MoveL 16 to (0, -3.6, 4.6) mm, rotated rx 0 ry 0 rz 180 deg; joints [18.023, -53.994, 108.608, -158.244, 56.588, 77.606]
  MoveL 17 to (0, -4.2, 4.6) mm, rotated rx 0 ry 0 rz 180 deg; joints [18.023, -54.022, 108.603, -158.236, 56.556, 77.591]
  MoveL 18 to (-200, -4.2, 4.6) mm, rotated rx 0 ry 0 rz 180 deg; joints [20.851, -62.892, 124.561, -156.601, 63.674, 79.137]
  MoveL 19 to (-200, -4.8, 4.6) mm, rotated rx 0 ry 0 rz 180 deg; joints [20.851, -62.926, 124.556, -156.593, 63.637, 79.119]
  MoveL 20 to (0, -4.8, 4.6) mm, rotated rx 0 ry 0 rz 180 deg; joints [18.023, -54.051, 108.598, -158.227, 56.525, 77.576]
  MoveL 21 to (0, -5.4, 4.6) mm, rotated rx 0 ry 0 rz 180 deg; joints [18.023, -54.08, 108.593, -158.219, 56.493, 77.561]
  MoveL 22 to (-200, -5.4, 4.6) mm, rotated rx 0 ry 0 rz 180 deg; joints [20.851, -62.961, 124.55, -156.585, 63.6, 79.101]
  MoveL 23 to (-200, -6, 4.6) mm, rotated rx 0 ry 0 rz 180 deg; joints [20.851, -62.996, 124.544, -156.577, 63.563, 79.083]
  MoveL 24 to (0, -6, 4.6) mm, rotated rx 0 ry 0 rz 180 deg; joints [18.023, -54.108, 108.588, -158.211, 56.462, 77.546]
  MoveL 25 to (0, -6.6, 4.6) mm, rotated rx 0 ry 0 rz 180 deg; joints [18.023, -54.137, 108.582, -158.202, 56.431, 77.531]
  MoveL 26 to (-200, -6.6, 4.6) mm, rotated rx 0 ry 0 rz 180 deg; joints [20.851, -63.031, 124.539, -156.569, 63.526, 79.065]
  MoveL 27 to (-200, -7.2, 4.6) mm, rotated rx 0 ry 0 rz 180 deg; joints [20.851, -63.066, 124.533, -156.561, 63.489, 79.047]
  MoveL 28 to (0, -7.2, 4.6) mm, rotated rx 0 ry 0 rz 180 deg; joints [18.023, -54.165, 108.577, -158.194, 56.399, 77.515]
  MoveL 29 to (0, -7.8, 4.6) mm, rotated rx 0 ry 0 rz 180 deg; joints [18.023, -54.194, 108.572, -158.186, 56.368, 77.5]
  MoveL 30 to (-200, -7.8, 4.6) mm, rotated rx 0 ry 0 rz 180 deg; joints [20.851, -63.1, 124.527, -156.553, 63.452, 79.029]
  MoveL 31 to (-200, -8.4, 4.6) mm, rotated rx 0 ry 0 rz 180 deg; joints [20.851, -63.135, 124.522, -156.545, 63.414, 79.011]
  MoveL 32 to (0, -8.4, 4.6) mm, rotated rx 0 ry 0 rz 180 deg; joints [18.023, -54.223, 108.567, -158.177, 56.336, 77.485]
  MoveL 33 to (0, -9, 4.6) mm, rotated rx 0 ry 0 rz 180 deg; joints [18.023, -54.251, 108.561, -158.169, 56.305, 77.47]
  MoveL 34 to (-200, -9, 4.6) mm, rotated rx 0 ry 0 rz 180 deg; joints [20.851, -63.17, 124.516, -156.537, 63.377, 78.993]
  MoveL 35 to (-200, -9.6, 4.6) mm, rotated rx 0 ry 0 rz 180 deg; joints [20.851, -63.204, 124.51, -156.529, 63.34, 78.975]
  MoveL 36 to (0, -9.6, 4.6) mm, rotated rx 0 ry 0 rz 180 deg; joints [18.023, -54.28, 108.556, -158.161, 56.273, 77.455]
  MoveL 37 to (0, -10.2, 4.6) mm, rotated rx 0 ry 0 rz 180 deg; joints [18.023, -54.308, 108.551, -158.152, 56.242, 77.44]
  MoveL 38 to (-200, -10.2, 4.6) mm, rotated rx 0 ry 0 rz 180 deg; joints [20.851, -63.239, 124.504, -156.521, 63.303, 78.957]
  MoveL 39 to (-200, -10.8, 4.6) mm, rotated rx 0 ry 0 rz 180 deg; joints [20.851, -63.274, 124.498, -156.513, 63.266, 78.939]
  MoveL 40 to (0, -10.8, 4.6) mm, rotated rx 0 ry 0 rz 180 deg; joints [18.023, -54.337, 108.545, -158.144, 56.211, 77.425]
  MoveL 41 to (0, -11.4, 4.6) mm, rotated rx 0 ry 0 rz 180 deg; joints [18.023, -54.365, 108.54, -158.135, 56.179, 77.409]
  MoveL 42 to (-200, -11.4, 4.6) mm, rotated rx 0 ry 0 rz 180 deg; joints [20.851, -63.308, 124.492, -156.505, 63.229, 78.921]
  MoveL 43 to (-200, -12, 4.6) mm, rotated rx 0 ry 0 rz 180 deg; joints [20.851, -63.343, 124.487, -156.497, 63.192, 78.903]
  MoveL 44 to (0, -12, 4.6) mm, rotated rx 0 ry 0 rz 180 deg; joints [18.023, -54.394, 108.534, -158.127, 56.148, 77.394]
  MoveL 45 to (0, -12.6, 4.6) mm, rotated rx 0 ry 0 rz 180 deg; joints [18.023, -54.422, 108.529, -158.118, 56.116, 77.379]
  MoveL 46 to (-200, -12.6, 4.6) mm, rotated rx 0 ry 0 rz 180 deg; joints [20.851, -63.378, 124.481, -156.488, 63.154, 78.885]
  MoveL 47 to (-200, -13.2, 4.6) mm, rotated rx 0 ry 0 rz 180 deg; joints [20.851, -63.412, 124.475, -156.48, 63.117, 78.867]
  MoveL 48 to (0, -13.2, 4.6) mm, rotated rx 0 ry 0 rz 180 deg; joints [18.023, -54.451, 108.523, -158.11, 56.085, 77.364]
  MoveL 49 to (0, -13.8, 4.6) mm, rotated rx 0 ry 0 rz 180 deg; joints [18.023, -54.479, 108.518, -158.101, 56.053, 77.348]
  MoveL 50 to (-200, -13.8, 4.6) mm, rotated rx 0 ry 0 rz 180 deg; joints [20.851, -63.447, 124.469, -156.472, 63.08, 78.849]
  MoveL 51 to (-200, -14.4, 4.6) mm, rotated rx 0 ry 0 rz 180 deg; joints [20.851, -63.481, 124.463, -156.464, 63.043, 78.83]
  MoveL 52 to (0, -14.4, 4.6) mm, rotated rx 0 ry 0 rz 180 deg; joints [18.023, -54.507, 108.512, -158.093, 56.021, 77.333]
  MoveL 53 to (0, -15, 4.6) mm, rotated rx 0 ry 0 rz 180 deg; joints [18.023, -54.536, 108.507, -158.084, 55.99, 77.318]
  MoveL 54 to (-200, -15, 4.6) mm, rotated rx 0 ry 0 rz 180 deg; joints [20.851, -63.516, 124.456, -156.455, 63.006, 78.812]
  MoveL 55 to (-200, -15.6, 4.6) mm, rotated rx 0 ry 0 rz 180 deg; joints [20.851, -63.55, 124.45, -156.447, 62.968, 78.794]
  MoveL 56 to (0, -15.6, 4.6) mm, rotated rx 0 ry 0 rz 180 deg; joints [18.023, -54.564, 108.501, -158.076, 55.958, 77.303]
  MoveL 57 to (0, -16.2, 4.6) mm, rotated rx 0 ry 0 rz 180 deg; joints [18.023, -54.593, 108.495, -158.067, 55.927, 77.287]
  MoveL 58 to (-200, -16.2, 4.6) mm, rotated rx 0 ry 0 rz 180 deg; joints [20.851, -63.585, 124.444, -156.439, 62.931, 78.776]
  MoveL 59 to (-200, -16.8, 4.6) mm, rotated rx 0 ry 0 rz 180 deg; joints [20.851, -63.619, 124.438, -156.431, 62.894, 78.758]
  MoveL 60 to (0, -16.8, 4.6) mm, rotated rx 0 ry 0 rz 180 deg; joints [18.023, -54.621, 108.49, -158.058, 55.895, 77.272]
  MoveL 61 to (0, -17.4, 4.6) mm, rotated rx 0 ry 0 rz 180 deg; joints [18.023, -54.649, 108.484, -158.05, 55.864, 77.256]
  MoveL 62 to (-200, -17.4, 4.6) mm, rotated rx 0 ry 0 rz 180 deg; joints [20.851, -63.653, 124.432, -156.422, 62.857, 78.739]
  MoveL 63 to (-200, -18, 4.6) mm, rotated rx 0 ry 0 rz 180 deg; joints [20.851, -63.688, 124.426, -156.414, 62.82, 78.721]
  MoveL 64 to (0, -18, 4.6) mm, rotated rx 0 ry 0 rz 180 deg; joints [18.023, -54.678, 108.478, -158.041, 55.832, 77.241]
  MoveL 65 to (0, -18.6, 4.6) mm, rotated rx 0 ry 0 rz 180 deg; joints [18.023, -54.706, 108.472, -158.032, 55.801, 77.226]
  MoveL 66 to (-200, -18.6, 4.6) mm, rotated rx 0 ry 0 rz 180 deg; joints [20.851, -63.722, 124.419, -156.406, 62.782, 78.703]
  MoveL 67 to (-200, -19.2, 4.6) mm, rotated rx 0 ry 0 rz 180 deg; joints [20.851, -63.756, 124.413, -156.397, 62.745, 78.685]
  MoveL 68 to (0, -19.2, 4.6) mm, rotated rx 0 ry 0 rz 180 deg; joints [18.023, -54.734, 108.466, -158.024, 55.769, 77.21]
  MoveL 69 to (0, -19.8, 4.6) mm, rotated rx 0 ry 0 rz 180 deg; joints [18.023, -54.762, 108.461, -158.015, 55.737, 77.195]
  MoveL 70 to (-200, -19.8, 4.6) mm, rotated rx 0 ry 0 rz 180 deg; joints [20.851, -63.791, 124.407, -156.389, 62.708, 78.666]
  MoveL 71 to (-200, -20.4, 4.6) mm, rotated rx 0 ry 0 rz 180 deg; joints [20.851, -63.825, 124.4, -156.38, 62.671, 78.648]
  MoveL 72 to (0, -20.4, 4.6) mm, rotated rx 0 ry 0 rz 180 deg; joints [18.023, -54.791, 108.455, -158.006, 55.706, 77.179]
  MoveL 73 to (0, -21, 4.6) mm, rotated rx 0 ry 0 rz 180 deg; joints [18.023, -54.819, 108.449, -157.998, 55.674, 77.164]
  MoveL 74 to (-200, -21, 4.6) mm, rotated rx 0 ry 0 rz 180 deg; joints [20.851, -63.859, 124.394, -156.372, 62.633, 78.63]
  MoveL 75 to (-200, -21.6, 4.6) mm, rotated rx 0 ry 0 rz 180 deg; joints [20.851, -63.894, 124.387, -156.364, 62.596, 78.611]
  MoveL 76 to (0, -21.6, 4.6) mm, rotated rx 0 ry 0 rz 180 deg; joints [18.023, -54.847, 108.443, -157.989, 55.642, 77.148]
  MoveL 77 to (0, -22.2, 4.6) mm, rotated rx 0 ry 0 rz 180 deg; joints [18.023, -54.875, 108.437, -157.98, 55.611, 77.133]
  MoveL 78 to (-200, -22.2, 4.6) mm, rotated rx 0 ry 0 rz 180 deg; joints [20.851, -63.928, 124.381, -156.355, 62.559, 78.593]
  MoveL 79 to (-200, -22.8, 4.6) mm, rotated rx 0 ry 0 rz 180 deg; joints [20.851, -63.962, 124.374, -156.347, 62.521, 78.574]
  MoveL 80 to (0, -22.8, 4.6) mm, rotated rx 0 ry 0 rz 180 deg; joints [18.023, -54.903, 108.431, -157.971, 55.579, 77.117]
  MoveL 81 to (0, -23.4, 4.6) mm, rotated rx 0 ry 0 rz 180 deg; joints [18.023, -54.931, 108.425, -157.963, 55.548, 77.102]
  MoveL 82 to (-200, -23.4, 4.6) mm, rotated rx 0 ry 0 rz 180 deg; joints [20.851, -63.996, 124.368, -156.338, 62.484, 78.556]
  MoveL 83 to (-200, -24, 4.6) mm, rotated rx 0 ry 0 rz 180 deg; joints [20.851, -64.03, 124.361, -156.33, 62.447, 78.538]
  MoveL 84 to (0, -24, 4.6) mm, rotated rx 0 ry 0 rz 180 deg; joints [18.023, -54.959, 108.419, -157.954, 55.516, 77.086]
  MoveL 85 to (0, -24.6, 4.6) mm, rotated rx 0 ry 0 rz 180 deg; joints [18.023, -54.988, 108.413, -157.945, 55.484, 77.071]
  MoveL 86 to (-200, -24.6, 4.6) mm, rotated rx 0 ry 0 rz 180 deg; joints [20.851, -64.065, 124.355, -156.321, 62.409, 78.519]
  MoveL 87 to (-200, -25.2, 4.6) mm, rotated rx 0 ry 0 rz 180 deg; joints [20.851, -64.099, 124.348, -156.312, 62.372, 78.501]
  MoveL 88 to (0, -25.2, 4.6) mm, rotated rx 0 ry 0 rz 180 deg; joints [18.023, -55.016, 108.407, -157.936, 55.453, 77.055]
  MoveL 89 to (0, -25.8, 4.6) mm, rotated rx 0 ry 0 rz 180 deg; joints [18.023, -55.044, 108.401, -157.927, 55.421, 77.04]
  MoveL 90 to (-200, -25.8, 4.6) mm, rotated rx 0 ry 0 rz 180 deg; joints [20.851, -64.133, 124.341, -156.304, 62.335, 78.482]
  MoveL 91 to (-200, -26.4, 4.6) mm, rotated rx 0 ry 0 rz 180 deg; joints [20.851, -64.167, 124.335, -156.295, 62.298, 78.464]
  MoveL 92 to (0, -26.4, 4.6) mm, rotated rx 0 ry 0 rz 180 deg; joints [18.023, -55.072, 108.394, -157.919, 55.389, 77.024]
  MoveL 93 to (0, -27, 4.6) mm, rotated rx 0 ry 0 rz 180 deg; joints [18.023, -55.1, 108.388, -157.91, 55.357, 77.008]
  MoveL 94 to (-200, -27, 4.6) mm, rotated rx 0 ry 0 rz 180 deg; joints [20.851, -64.201, 124.328, -156.287, 62.26, 78.445]
  MoveL 95 to (-200, -27.6, 4.6) mm, rotated rx 0 ry 0 rz 180 deg; joints [20.851, -64.235, 124.321, -156.278, 62.223, 78.427]
  MoveL 96 to (0, -27.6, 4.6) mm, rotated rx 0 ry 0 rz 180 deg; joints [18.023, -55.128, 108.382, -157.901, 55.326, 76.993]
  MoveL 97 to (0, -28.2, 4.6) mm, rotated rx 0 ry 0 rz 180 deg; joints [18.023, -55.156, 108.376, -157.892, 55.294, 76.977]
  MoveL 98 to (-200, -28.2, 4.6) mm, rotated rx 0 ry 0 rz 180 deg; joints [20.851, -64.269, 124.314, -156.269, 62.185, 78.408]
  MoveL 99 to (-200, -28.8, 4.6) mm, rotated rx 0 ry 0 rz 180 deg; joints [20.851, -64.303, 124.308, -156.261, 62.148, 78.389]
  MoveL 100 to (0, -28.8, 4.6) mm, rotated rx 0 ry 0 rz 180 deg; joints [18.023, -55.184, 108.37, -157.883, 55.262, 76.961]
  MoveL 101 to (0, -29.4, 4.6) mm, rotated rx 0 ry 0 rz 180 deg; joints [18.023, -55.212, 108.363, -157.874, 55.231, 76.946]
  MoveL 102 to (-200, -29.4, 4.6) mm, rotated rx 0 ry 0 rz 180 deg; joints [20.851, -64.337, 124.301, -156.252, 62.111, 78.371]
  MoveL 103 to (-200, -30, 4.6) mm, rotated rx 0 ry 0 rz 180 deg; joints [20.851, -64.371, 124.294, -156.243, 62.073, 78.352]
  MoveL 104 to (0, -30, 4.6) mm, rotated rx 0 ry 0 rz 180 deg; joints [18.023, -55.24, 108.357, -157.865, 55.199, 76.93]
  MoveL 105 to (0, -30.6, 4.62) mm, rotated rx 3.31 ry 0 rz 180 deg; joints [17.906, -56.261, 108.2, -157.689, 54.081, 79.771]
  MoveL 106 to (-200, -30.6, 4.62) mm, rotated rx 3.31 ry 0 rz 180 deg; joints [20.718, -65.607, 124.119, -156.08, 60.756, 81.08]
  MoveL 107 to (-200, -31.2, 4.67) mm, rotated rx 6.61 ry 0 rz 180 deg; joints [20.534, -66.826, 123.942, -155.962, 59.439, 83.834]
  MoveL 108 to (0, -31.2, 4.67) mm, rotated rx 6.61 ry 0 rz 180 deg; joints [17.742, -57.27, 108.042, -157.558, 52.964, 82.641]
  MoveL 109 to (0, -31.79, 4.75) mm, rotated rx 9.92 ry 0 rz 180 deg; joints [17.533, -58.264, 107.884, -157.475, 51.848, 85.547]
  MoveL 110 to (-200, -31.79, 4.75) mm, rotated rx 9.92 ry 0 rz 180 deg; joints [20.297, -68.026, 123.763, -155.891, 58.127, 86.622]
  MoveL 111 to (-200, -32.38, 4.88) mm, rotated rx 13.22 ry 0 rz 180 deg; joints [20.008, -69.203, 123.584, -155.871, 56.821, 89.448]
  MoveL 112 to (0, -32.38, 4.88) mm, rotated rx 13.22 ry 0 rz 180 deg; joints [17.278, -59.239, 107.727, -157.443, 50.738, 88.493]
  MoveL 113 to (0, -32.96, 5.03) mm, rotated rx 16.53 ry 0 rz 180 deg; joints [16.978, -60.194, 107.571, -157.465, 49.635, 91.486]
  MoveL 114 to (-200, -32.96, 5.03) mm, rotated rx 16.53 ry 0 rz 180 deg; joints [19.668, -70.354, 123.404, -155.904, 55.525, 92.321]
  MoveL 115 to (-200, -33.53, 5.22) mm, rotated rx 19.83 ry 0 rz 180 deg; joints [19.277, -71.476, 123.226, -155.994, 54.241, 95.245]
  MoveL 116 to (0, -33.53, 5.22) mm, rotated rx 19.83 ry 0 rz 180 deg; joints [16.634, -61.125, 107.418, -157.545, 48.543, 94.53]
  MoveL 117 to (0, -34.09, 5.44) mm, rotated rx 23.14 ry 0 rz 180 deg; joints [16.246, -62.031, 107.268, -157.686, 47.464, 97.632]
  MoveL 118 to (-200, -34.09, 5.44) mm, rotated rx 23.14 ry 0 rz 180 deg; joints [18.836, -72.566, 123.051, -156.146, 52.973, 98.228]
  MoveL 119 to (-200, -34.63, 5.69) mm, rotated rx 26.44 ry 0 rz 180 deg; joints [18.346, -73.62, 122.881, -156.363, 51.724, 101.275]
  MoveL 120 to (0, -34.63, 5.69) mm, rotated rx 26.44 ry 0 rz 180 deg; joints [15.816, -62.908, 107.123, -157.893, 46.402, 100.796]
  MoveL 121 to (0, -35.16, 5.97) mm, rotated rx 29.75 ry 0 rz 180 deg; joints [15.343, -63.755, 106.984, -158.169, 45.36, 104.029]
  MoveL 122 to (-200, -35.16, 5.97) mm, rotated rx 29.75 ry 0 rz 180 deg; joints [17.807, -74.638, 122.715, -156.651, 50.497, 104.395]
  MoveL 123 to (-200, -35.67, 6.28) mm, rotated rx 33.05 ry 0 rz 180 deg; joints [17.221, -75.615, 122.557, -157.013, 49.297, 107.592]
  MoveL 124 to (0, -35.67, 6.28) mm, rotated rx 33.05 ry 0 rz 180 deg; joints [14.829, -64.568, 106.852, -158.519, 44.342, 107.336]
  MoveL 125 to (0, -36.17, 6.62) mm, rotated rx 36.36 ry 0 rz 180 deg; joints [14.276, -65.347, 106.728, -158.947, 43.351, 110.724]
  MoveL 126 to (-200, -36.17, 6.62) mm, rotated rx 36.36 ry 0 rz 180 deg; joints [16.588, -76.55, 122.407, -157.456, 48.127, 110.874]
  MoveL 127 to (-200, -36.64, 6.99) mm, rotated rx 39.67 ry 0 rz 180 deg; joints [15.91, -77.44, 122.266, -157.984, 46.993, 114.247]
  MoveL 128 to (0, -36.64, 6.99) mm, rotated rx 39.67 ry 0 rz 180 deg; joints [13.685, -66.088, 106.614, -159.457, 42.393, 114.196]
  MoveL 129 to (0, -37.09, 7.39) mm, rotated rx 42.97 ry 0 rz 180 deg; joints [13.057, -66.79, 106.51, -160.053, 41.47, 117.759]
  MoveL 130 to (-200, -37.09, 7.39) mm, rotated rx 42.97 ry 0 rz 180 deg; joints [15.189, -78.283, 122.137, -158.602, 45.899, 117.718]
  MoveL 131 to (-200, -37.52, 7.81) mm, rotated rx 46.28 ry 0 rz 180 deg; joints [14.427, -79.077, 122.02, -159.313, 44.851, 121.29]
  MoveL 132 to (0, -37.52, 7.81) mm, rotated rx 46.28 ry 0 rz 180 deg; joints [12.394, -67.452, 106.418, -160.738, 40.589, 121.415]
  MoveL 133 to (0, -37.92, 8.26) mm, rotated rx 49.58 ry 0 rz 180 deg; joints [11.697, -68.07, 106.338, -161.515, 39.752, 125.169]
  MoveL 134 to (-200, -37.92, 8.26) mm, rotated rx 49.58 ry 0 rz 180 deg; joints [13.624, -79.819, 121.917, -160.123, 43.853, 124.971]
  MoveL 135 to (-200, -38.29, 8.72) mm, rotated rx 52.89 ry 0 rz 180 deg; joints [12.785, -80.507, 121.829, -161.034, 42.913, 128.76]
  MoveL 136 to (0, -38.29, 8.72) mm, rotated rx 52.89 ry 0 rz 180 deg; joints [10.97, -68.644, 106.272, -162.386, 38.967, 129.022]
  MoveL 137 to (0, -38.64, 9.21) mm, rotated rx 56.19 ry 0 rz 180 deg; joints [10.214, -69.171, 106.222, -163.351, 38.237, 132.976]
  MoveL 138 to (-200, -38.64, 9.21) mm, rotated rx 56.19 ry 0 rz 180 deg; joints [11.911, -81.141, 121.757, -162.047, 42.035, 132.663]
  MoveL 139 to (-200, -38.96, 9.72) mm, rotated rx 59.5 ry 0 rz 180 deg; joints [11.005, -81.717, 121.703, -163.163, 41.226, 136.677]
  MoveL 140 to (0, -38.96, 9.72) mm, rotated rx 59.5 ry 0 rz 180 deg; joints [9.432, -69.651, 106.186, -164.409, 37.568, 137.028]
  MoveL 141 to (0, -39.25, 10.25) mm, rotated rx 62.8 ry 0 rz 180 deg; joints [8.625, -70.082, 106.167, -165.559, 36.965, 141.178]
  MoveL 142 to (-200, -39.25, 10.25) mm, rotated rx 62.8 ry 0 rz 180 deg; joints [10.069, -82.235, 121.667, -164.381, 40.494, 140.803]
  MoveL 143 to (-200, -39.51, 10.79) mm, rotated rx 66.11 ry 0 rz 180 deg; joints [9.107, -82.692, 121.651, -165.697, 39.843, 145.035]
  MoveL 144 to (0, -39.51, 10.79) mm, rotated rx 66.11 ry 0 rz 180 deg; joints [7.797, -70.462, 106.166, -166.795, 36.434, 145.421]
  MoveL 145 to (0, -39.74, 11.34) mm, rotated rx 69.42 ry 0 rz 180 deg; joints [6.951, -70.791, 106.181, -168.111, 35.979, 149.748]
  MoveL 146 to (-200, -39.74, 11.34) mm, rotated rx 69.42 ry 0 rz 180 deg; joints [8.123, -83.088, 121.654, -167.105, 39.282, 149.367]
  MoveL 147 to (-200, -39.93, 11.91) mm, rotated rx 72.72 ry 0 rz 180 deg; joints [7.119, -83.421, 121.678, -168.596, 38.814, 153.79]
  MoveL 148 to (0, -39.93, 11.91) mm, rotated rx 72.72 ry 0 rz 180 deg; joints [6.09, -71.068, 106.215, -169.5, 35.604, 154.153]
  MoveL 149 to (0, -40.09, 12.49) mm, rotated rx 76.03 ry 0 rz 180 deg; joints [5.217, -71.291, 106.267, -170.95, 35.314, 158.622]
  MoveL 150 to (-200, -40.09, 12.49) mm, rotated rx 76.03 ry 0 rz 180 deg; joints [6.101, -83.69, 121.723, -170.158, 38.446, 158.29]
  MoveL 151 to (-200, -40.22, 13.07) mm, rotated rx 79.33 ry 0 rz 180 deg; joints [5.071, -83.894, 121.79, -171.78, 38.183, 162.855]
  MoveL 152 to (0, -40.22, 13.07) mm, rotated rx 79.33 ry 0 rz 180 deg; joints [4.334, -71.46, 106.338, -172.45, 35.112, 163.145]
  MoveL 153 to (0, -40.31, 13.67) mm, rotated rx 82.64 ry 0 rz 180 deg; joints [3.447, -71.574, 106.427, -173.984, 35.002, 167.704]
  MoveL 154 to (-200, -40.31, 13.67) mm, rotated rx 82.64 ry 0 rz 180 deg; joints [4.033, -84.032, 121.877, -173.444, 38.027, 167.465]
  MoveL 155 to (-200, -40.37, 14.26) mm, rotated rx 85.94 ry 0 rz 180 deg; joints [2.992, -84.104, 121.986, -175.135, 37.983, 172.106]
  MoveL 156 to (0, -40.37, 14.26) mm, rotated rx 85.94 ry 0 rz 180 deg; joints [2.556, -71.632, 106.534, -175.538, 34.983, 172.286]
  MoveL 157 to (0, -40.4, 14.86) mm, rotated rx 89.25 ry 0 rz 180 deg; joints [1.668, -71.635, 106.659, -177.096, 35.059, 176.871]
  MoveL 158 to (-200, -40.4, 14.86) mm, rotated rx 89.25 ry 0 rz 180 deg; joints [1.952, -84.108, 122.116, -176.832, 38.05, 176.753]
  MoveL 159 to (-200, -40.4, 15.46) mm, rotated rx 90 ry 0 rz 180 deg; joints [1.693, -84.101, 122.149, -177.254, 38.08, 177.838]
  MoveL 160 to (0, -40.4, 15.46) mm, rotated rx 90 ry 0 rz 180 deg; joints [1.447, -71.628, 106.69, -177.483, 35.088, 177.94]
  MoveL 161 to (0, -40.4, 16.06) mm, rotated rx 90 ry 0 rz 180 deg; joints [1.422, -71.629, 106.692, -177.526, 35.088, 177.975]
  MoveL 162 to (-200, -40.4, 16.06) mm, rotated rx 90 ry 0 rz 180 deg; joints [1.664, -84.102, 122.15, -177.301, 38.079, 177.875]
  MoveL 163 to (-200, -40.4, 16.66) mm, rotated rx 90 ry 0 rz 180 deg; joints [1.635, -84.103, 122.152, -177.349, 38.078, 177.912]
  MoveL 164 to (0, -40.4, 16.66) mm, rotated rx 90 ry 0 rz 180 deg; joints [1.397, -71.63, 106.693, -177.57, 35.087, 178.011]
  MoveL 165 to (0, -40.4, 17.26) mm, rotated rx 90 ry 0 rz 180 deg; joints [1.372, -71.631, 106.694, -177.613, 35.087, 178.047]
  MoveL 166 to (-200, -40.4, 17.26) mm, rotated rx 90 ry 0 rz 180 deg; joints [1.606, -84.104, 122.153, -177.396, 38.077, 177.95]
  MoveL 167 to (-200, -40.4, 17.86) mm, rotated rx 90 ry 0 rz 180 deg; joints [1.576, -84.105, 122.154, -177.444, 38.076, 177.987]
  MoveL 168 to (0, -40.4, 17.86) mm, rotated rx 90 ry 0 rz 180 deg; joints [1.347, -71.632, 106.695, -177.657, 35.086, 178.082]
  MoveL 169 to (0, -40.4, 18.46) mm, rotated rx 90 ry 0 rz 180 deg; joints [1.321, -71.632, 106.696, -177.701, 35.086, 178.118]
  MoveL 170 to (-200, -40.4, 18.46) mm, rotated rx 90 ry 0 rz 180 deg; joints [1.547, -84.106, 122.155, -177.491, 38.076, 178.025]
  MoveL 171 to (-200, -40.4, 19.06) mm, rotated rx 90 ry 0 rz 180 deg; joints [1.518, -84.107, 122.156, -177.539, 38.075, 178.062]
  MoveL 172 to (0, -40.4, 19.06) mm, rotated rx 90 ry 0 rz 180 deg; joints [1.296, -71.633, 106.698, -177.744, 35.085, 178.154]
  MoveL 173 to (0, -40.4, 19.66) mm, rotated rx 90 ry 0 rz 180 deg; joints [1.271, -71.634, 106.699, -177.788, 35.085, 178.189]
  MoveL 174 to (-200, -40.4, 19.66) mm, rotated rx 90 ry 0 rz 180 deg; joints [1.488, -84.108, 122.157, -177.586, 38.074, 178.099]
  MoveL 175 to (-200, -40.4, 20.26) mm, rotated rx 90 ry 0 rz 180 deg; joints [1.459, -84.109, 122.159, -177.634, 38.073, 178.137]
  MoveL 176 to (0, -40.4, 20.26) mm, rotated rx 90 ry 0 rz 180 deg; joints [1.246, -71.635, 106.7, -177.831, 35.084, 178.225]
  MoveL 177 to (0, -40.4, 20.86) mm, rotated rx 90 ry 0 rz 180 deg; joints [1.221, -71.636, 106.701, -177.875, 35.084, 178.261]
  MoveL 178 to (-200, -40.4, 20.86) mm, rotated rx 90 ry 0 rz 180 deg; joints [1.43, -84.11, 122.16, -177.681, 38.072, 178.174]
  MoveL 179 to (-200, -40.4, 21.46) mm, rotated rx 90 ry 0 rz 180 deg; joints [1.4, -84.111, 122.161, -177.729, 38.071, 178.212]
  MoveL 180 to (0, -40.4, 21.46) mm, rotated rx 90 ry 0 rz 180 deg; joints [1.196, -71.637, 106.702, -177.918, 35.083, 178.296]
  MoveL 181 to (0, -40.4, 22.06) mm, rotated rx 90 ry 0 rz 180 deg; joints [1.171, -71.637, 106.703, -177.962, 35.083, 178.332]
  MoveL 182 to (-200, -40.4, 22.06) mm, rotated rx 90 ry 0 rz 180 deg; joints [1.371, -84.112, 122.162, -177.776, 38.071, 178.249]
  MoveL 183 to (-200, -40.4, 22.66) mm, rotated rx 90 ry 0 rz 180 deg; joints [1.342, -84.113, 122.163, -177.824, 38.07, 178.286]
  MoveL 184 to (0, -40.4, 22.66) mm, rotated rx 90 ry 0 rz 180 deg; joints [1.146, -71.638, 106.704, -178.006, 35.082, 178.368]
  MoveL 185 to (0, -40.4, 23.26) mm, rotated rx 90 ry 0 rz 180 deg; joints [1.121, -71.639, 106.705, -178.049, 35.082, 178.403]
  MoveL 186 to (-200, -40.4, 23.26) mm, rotated rx 90 ry 0 rz 180 deg; joints [1.312, -84.114, 122.164, -177.871, 38.069, 178.324]
  MoveL 187 to (-200, -40.4, 23.86) mm, rotated rx 90 ry 0 rz 180 deg; joints [1.283, -84.115, 122.165, -177.919, 38.068, 178.361]
  MoveL 188 to (0, -40.4, 23.86) mm, rotated rx 90 ry 0 rz 180 deg; joints [1.096, -71.639, 106.706, -178.093, 35.081, 178.439]
  MoveL 189 to (0, -40.4, 24.46) mm, rotated rx 90 ry 0 rz 180 deg; joints [1.071, -71.64, 106.707, -178.136, 35.081, 178.475]
  MoveL 190 to (-200, -40.4, 24.46) mm, rotated rx 90 ry 0 rz 180 deg; joints [1.254, -84.116, 122.166, -177.966, 38.068, 178.399]
  MoveL 191 to (-200, -40.4, 25.06) mm, rotated rx 90 ry 0 rz 180 deg; joints [1.224, -84.117, 122.167, -178.014, 38.067, 178.436]
  MoveL 192 to (0, -40.4, 25.06) mm, rotated rx 90 ry 0 rz 180 deg; joints [1.046, -71.641, 106.708, -178.18, 35.08, 178.51]
  MoveL 193 to (0, -40.4, 25.66) mm, rotated rx 90 ry 0 rz 180 deg; joints [1.021, -71.642, 106.709, -178.223, 35.08, 178.546]
  MoveL 194 to (-200, -40.4, 25.66) mm, rotated rx 90 ry 0 rz 180 deg; joints [1.195, -84.117, 122.168, -178.061, 38.066, 178.474]
  MoveL 195 to (-200, -40.4, 26.26) mm, rotated rx 90 ry 0 rz 180 deg; joints [1.166, -84.118, 122.168, -178.109, 38.065, 178.511]
  MoveL 196 to (0, -40.4, 26.26) mm, rotated rx 90 ry 0 rz 180 deg; joints [0.996, -71.642, 106.71, -178.267, 35.08, 178.582]
  MoveL 197 to (0, -40.4, 26.86) mm, rotated rx 90 ry 0 rz 180 deg; joints [0.971, -71.643, 106.71, -178.311, 35.079, 178.617]
  MoveL 198 to (-200, -40.4, 26.86) mm, rotated rx 90 ry 0 rz 180 deg; joints [1.136, -84.119, 122.169, -178.157, 38.065, 178.548]
  MoveL 199 to (-200, -40.4, 27.46) mm, rotated rx 90 ry 0 rz 180 deg; joints [1.107, -84.12, 122.17, -178.204, 38.064, 178.586]
  MoveL 200 to (0, -40.4, 27.46) mm, rotated rx 90 ry 0 rz 180 deg; joints [0.946, -71.643, 106.711, -178.354, 35.079, 178.653]
  MoveL 201 to (0, -40.4, 28.06) mm, rotated rx 90 ry 0 rz 180 deg; joints [0.921, -71.644, 106.712, -178.398, 35.079, 178.689]
  MoveL 202 to (-200, -40.4, 28.06) mm, rotated rx 90 ry 0 rz 180 deg; joints [1.078, -84.12, 122.171, -178.252, 38.063, 178.623]
  MoveL 203 to (-200, -40.4, 28.66) mm, rotated rx 90 ry 0 rz 180 deg; joints [1.048, -84.121, 122.172, -178.299, 38.063, 178.661]
  MoveL 204 to (0, -40.4, 28.66) mm, rotated rx 90 ry 0 rz 180 deg; joints [0.896, -71.645, 106.713, -178.441, 35.078, 178.724]
  MoveL 205 to (0, -40.4, 29.26) mm, rotated rx 90 ry 0 rz 180 deg; joints [0.871, -71.645, 106.714, -178.485, 35.078, 178.76]
  MoveL 206 to (-200, -40.4, 29.26) mm, rotated rx 90 ry 0 rz 180 deg; joints [1.019, -84.122, 122.173, -178.347, 38.062, 178.698]
  MoveL 207 to (-200, -40.4, 29.86) mm, rotated rx 90 ry 0 rz 180 deg; joints [0.99, -84.122, 122.173, -178.394, 38.062, 178.736]
  MoveL 208 to (0, -40.4, 29.86) mm, rotated rx 90 ry 0 rz 180 deg; joints [0.846, -71.646, 106.714, -178.529, 35.078, 178.796]
  MoveL 209 to (0, -40.4, 30.46) mm, rotated rx 90 ry 0 rz 180 deg; joints [0.821, -71.646, 106.715, -178.572, 35.077, 178.831]
  MoveL 210 to (-200, -40.4, 30.46) mm, rotated rx 90 ry 0 rz 180 deg; joints [0.961, -84.123, 122.174, -178.442, 38.061, 178.773]
  MoveL 211 to (-200, -40.4, 31.06) mm, rotated rx 90 ry 0 rz 180 deg; joints [0.931, -84.124, 122.175, -178.489, 38.061, 178.811]
  MoveL 212 to (0, -40.4, 31.06) mm, rotated rx 90 ry 0 rz 180 deg; joints [0.795, -71.647, 106.716, -178.616, 35.077, 178.867]
  MoveL 213 to (0, -40.4, 31.66) mm, rotated rx 90 ry 0 rz 180 deg; joints [0.77, -71.647, 106.716, -178.659, 35.077, 178.903]
  MoveL 214 to (-200, -40.4, 31.66) mm, rotated rx 90 ry 0 rz 180 deg; joints [0.902, -84.124, 122.175, -178.537, 38.06, 178.848]
  MoveL 215 to (-200, -40.4, 32.26) mm, rotated rx 90 ry 0 rz 180 deg; joints [0.873, -84.125, 122.176, -178.585, 38.06, 178.885]
  MoveL 216 to (0, -40.4, 32.26) mm, rotated rx 90 ry 0 rz 180 deg; joints [0.745, -71.648, 106.717, -178.703, 35.076, 178.938]
  MoveL 217 to (0, -40.4, 32.86) mm, rotated rx 90 ry 0 rz 180 deg; joints [0.72, -71.648, 106.718, -178.746, 35.076, 178.974]
  MoveL 218 to (-200, -40.4, 32.86) mm, rotated rx 90 ry 0 rz 180 deg; joints [0.843, -84.126, 122.177, -178.632, 38.059, 178.923]
  MoveL 219 to (-200, -40.4, 33.46) mm, rotated rx 90 ry 0 rz 180 deg; joints [0.814, -84.126, 122.177, -178.68, 38.059, 178.96]
  MoveL 220 to (0, -40.4, 33.46) mm, rotated rx 90 ry 0 rz 180 deg; joints [0.695, -71.649, 106.718, -178.79, 35.076, 179.01]
  MoveL 221 to (0, -40.4, 34.06) mm, rotated rx 90 ry 0 rz 180 deg; joints [0.67, -71.649, 106.719, -178.834, 35.075, 179.045]
  MoveL 222 to (-200, -40.4, 34.06) mm, rotated rx 90 ry 0 rz 180 deg; joints [0.785, -84.127, 122.178, -178.727, 38.058, 178.998]
  MoveL 223 to (-200, -40.4, 34.66) mm, rotated rx 90 ry 0 rz 180 deg; joints [0.755, -84.127, 122.179, -178.775, 38.058, 179.035]
  MoveL 224 to (0, -40.4, 34.66) mm, rotated rx 90 ry 0 rz 180 deg; joints [0.645, -71.65, 106.72, -178.877, 35.075, 179.081]
  MoveL 225 to (0, -40.4, 35.26) mm, rotated rx 90 ry 0 rz 180 deg; joints [0.62, -71.65, 106.72, -178.921, 35.075, 179.117]
  MoveL 226 to (-200, -40.4, 35.26) mm, rotated rx 90 ry 0 rz 180 deg; joints [0.726, -84.128, 122.179, -178.822, 38.057, 179.073]
  MoveL 227 to (-200, -40.4, 35.86) mm, rotated rx 90 ry 0 rz 180 deg; joints [0.697, -84.128, 122.18, -178.87, 38.057, 179.11]
  MoveL 228 to (0, -40.4, 35.86) mm, rotated rx 90 ry 0 rz 180 deg; joints [0.595, -71.65, 106.721, -178.964, 35.075, 179.152]
  MoveL 229 to (0, -40.4, 36.46) mm, rotated rx 90 ry 0 rz 180 deg; joints [0.57, -71.651, 106.721, -179.008, 35.074, 179.188]
  MoveL 230 to (-200, -40.4, 36.46) mm, rotated rx 90 ry 0 rz 180 deg; joints [0.667, -84.129, 122.18, -178.918, 38.056, 179.148]
  MoveL 231 to (-200, -40.4, 37.06) mm, rotated rx 90 ry 0 rz 180 deg; joints [0.638, -84.129, 122.181, -178.965, 38.056, 179.185]
  MoveL 232 to (0, -40.4, 37.06) mm, rotated rx 90 ry 0 rz 180 deg; joints [0.545, -71.651, 106.722, -179.052, 35.074, 179.224]
  MoveL 233 to (0, -40.4, 37.66) mm, rotated rx 90 ry 0 rz 180 deg; joints [0.52, -71.651, 106.722, -179.095, 35.074, 179.26]
  MoveL 234 to (-200, -40.4, 37.66) mm, rotated rx 90 ry 0 rz 180 deg; joints [0.609, -84.129, 122.181, -179.013, 38.056, 179.223]
  MoveL 235 to (-200, -40.4, 38.26) mm, rotated rx 90 ry 0 rz 180 deg; joints [0.579, -84.13, 122.182, -179.06, 38.055, 179.26]
  MoveL 236 to (0, -40.4, 38.26) mm, rotated rx 90 ry 0 rz 180 deg; joints [0.495, -71.652, 106.723, -179.139, 35.074, 179.295]
  MoveL 237 to (0, -40.4, 38.86) mm, rotated rx 90 ry 0 rz 180 deg; joints [0.47, -71.652, 106.723, -179.182, 35.074, 179.331]
  MoveL 238 to (-200, -40.4, 38.86) mm, rotated rx 90 ry 0 rz 180 deg; joints [0.55, -84.13, 122.182, -179.108, 38.055, 179.297]
  MoveL 239 to (-200, -40.4, 39.46) mm, rotated rx 90 ry 0 rz 180 deg; joints [0.521, -84.131, 122.182, -179.155, 38.055, 179.335]
  MoveL 240 to (0, -40.4, 39.46) mm, rotated rx 90 ry 0 rz 180 deg; joints [0.445, -71.652, 106.723, -179.226, 35.073, 179.367]
  MoveL 241 to (0, -40.4, 40.06) mm, rotated rx 90 ry 0 rz 180 deg; joints [0.42, -71.653, 106.724, -179.27, 35.073, 179.402]
  MoveL 242 to (-200, -40.4, 40.06) mm, rotated rx 90 ry 0 rz 180 deg; joints [0.491, -84.131, 122.183, -179.203, 38.054, 179.372]
  MoveL 243 to (-200, -40.4, 40.66) mm, rotated rx 90 ry 0 rz 180 deg; joints [0.462, -84.131, 122.183, -179.251, 38.054, 179.41]
  MoveL 244 to (0, -40.4, 40.66) mm, rotated rx 90 ry 0 rz 180 deg; joints [0.395, -71.653, 106.724, -179.313, 35.073, 179.438]
  MoveL 245 to (0, -40.4, 41.26) mm, rotated rx 90 ry 0 rz 180 deg; joints [0.37, -71.653, 106.724, -179.357, 35.073, 179.474]
  MoveL 246 to (-200, -40.4, 41.26) mm, rotated rx 90 ry 0 rz 180 deg; joints [0.433, -84.132, 122.183, -179.298, 38.054, 179.447]
  MoveL 247 to (-200, -40.4, 41.86) mm, rotated rx 90 ry 0 rz 180 deg; joints [0.403, -84.132, 122.184, -179.346, 38.054, 179.485]
  MoveL 248 to (0, -40.4, 41.86) mm, rotated rx 90 ry 0 rz 180 deg; joints [0.344, -71.653, 106.725, -179.4, 35.073, 179.509]
  MoveL 249 to (0, -40.4, 42.46) mm, rotated rx 90 ry 0 rz 180 deg; joints [0.319, -71.654, 106.725, -179.444, 35.073, 179.545]
  MoveL 250 to (-200, -40.4, 42.46) mm, rotated rx 90 ry 0 rz 180 deg; joints [0.374, -84.132, 122.184, -179.393, 38.053, 179.522]
  MoveL 251 to (-200, -40.4, 43.06) mm, rotated rx 90 ry 0 rz 180 deg; joints [0.345, -84.132, 122.184, -179.441, 38.053, 179.56]
  MoveL 252 to (0, -40.4, 43.06) mm, rotated rx 90 ry 0 rz 180 deg; joints [0.294, -71.654, 106.725, -179.488, 35.073, 179.581]
  MoveL 253 to (0, -40.4, 43.66) mm, rotated rx 90 ry 0 rz 180 deg; joints [0.269, -71.654, 106.726, -179.531, 35.072, 179.616]
  MoveL 254 to (-200, -40.4, 43.66) mm, rotated rx 90 ry 0 rz 180 deg; joints [0.315, -84.133, 122.185, -179.489, 38.053, 179.597]
  MoveL 255 to (-200, -40.4, 44.26) mm, rotated rx 90 ry 0 rz 180 deg; joints [0.286, -84.133, 122.185, -179.536, 38.053, 179.635]
  MoveL 256 to (0, -40.4, 44.26) mm, rotated rx 90 ry 0 rz 180 deg; joints [0.244, -71.654, 106.726, -179.575, 35.072, 179.652]
  MoveL 257 to (0, -40.4, 44.86) mm, rotated rx 90 ry 0 rz 180 deg; joints [0.219, -71.654, 106.726, -179.619, 35.072, 179.688]
  MoveL 258 to (-200, -40.4, 44.86) mm, rotated rx 90 ry 0 rz 180 deg; joints [0.257, -84.133, 122.185, -179.584, 38.053, 179.672]
  MoveL 259 to (-200, -40.39, 45.46) mm, rotated rx 92.55 ry 0 rz 180 deg; joints [-0.55, -84.052, 122.273, 179.111, 38.224, -176.747]
  MoveL 260 to (0, -40.39, 45.46) mm, rotated rx 92.55 ry 0 rz 180 deg; joints [-0.47, -71.586, 106.808, 179.185, 35.224, -176.779]
  MoveL 261 to (0, -40.35, 46.06) mm, rotated rx 95.86 ry 0 rz 180 deg; joints [-1.346, -71.448, 106.928, 177.682, 35.502, -172.252]
  MoveL 262 to (-200, -40.35, 46.06) mm, rotated rx 95.86 ry 0 rz 180 deg; joints [-1.576, -83.887, 122.404, 177.471, 38.544, -172.161]
  MoveL 263 to (-200, -40.27, 46.66) mm, rotated rx 99.17 ry 0 rz 180 deg; joints [-2.588, -83.655, 122.554, 175.883, 38.972, -167.631]
  MoveL 264 to (0, -40.27, 46.66) mm, rotated rx 99.17 ry 0 rz 180 deg; joints [-2.211, -71.255, 107.065, 176.225, 35.869, -167.773]
  MoveL 265 to (0, -40.16, 47.25) mm, rotated rx 102.47 ry 0 rz 180 deg; joints [-3.06, -71.006, 107.218, 174.829, 36.323, -163.359]
  MoveL 266 to (-200, -40.16, 47.25) mm, rotated rx 102.47 ry 0 rz 180 deg; joints [-3.581, -83.357, 122.723, 174.365, 39.503, -163.175]
  MoveL 267 to (-200, -40.01, 47.83) mm, rotated rx 105.78 ry 0 rz 180 deg; joints [-4.553, -82.992, 122.909, 172.925, 40.133, -158.803]
  MoveL 268 to (0, -40.01, 47.83) mm, rotated rx 105.78 ry 0 rz 180 deg; joints [-3.892, -70.703, 107.384, 173.503, 36.859, -159.017]
  MoveL 269 to (0, -39.83, 48.4) mm, rotated rx 109.08 ry 0 rz 180 deg; joints [-4.702, -70.345, 107.565, 172.257, 37.473, -154.759]
  MoveL 270 to (-200, -39.83, 48.4) mm, rotated rx 109.08 ry 0 rz 180 deg; joints [-5.5, -82.562, 123.111, 171.575, 40.856, -154.526]
  MoveL 271 to (-200, -39.62, 48.96) mm, rotated rx 112.39 ry 0 rz 180 deg; joints [-6.417, -82.067, 123.327, 170.321, 41.667, -150.351]
  MoveL 272 to (0, -39.62, 48.96) mm, rotated rx 112.39 ry 0 rz 180 deg; joints [-5.488, -69.934, 107.757, 171.095, 38.16, -150.589]
  MoveL 273 to (0, -39.37, 49.51) mm, rotated rx 115.69 ry 0 rz 180 deg; joints [-6.247, -69.471, 107.96, 170.024, 38.915, -146.514]
  MoveL 274 to (-200, -39.37, 49.51) mm, rotated rx 115.69 ry 0 rz 180 deg; joints [-7.303, -81.509, 123.556, 169.168, 42.56, -146.285]
  MoveL 275 to (-200, -39.1, 50.04) mm, rotated rx 119 ry 0 rz 180 deg; joints [-8.153, -80.889, 123.797, 168.116, 43.527, -142.326]
  MoveL 276 to (0, -39.1, 50.04) mm, rotated rx 119 ry 0 rz 180 deg; joints [-6.977, -68.957, 108.173, 169.045, 39.734, -142.534]
  MoveL 277 to (0, -38.79, 50.56) mm, rotated rx 122.3 ry 0 rz 180 deg; joints [-7.675, -68.392, 108.394, 168.159, 40.609, -138.653]
  MoveL 278 to (-200, -38.79, 50.56) mm, rotated rx 122.3 ry 0 rz 180 deg; joints [-8.965, -80.208, 124.047, 167.168, 44.563, -138.478]
  MoveL 279 to (-200, -38.45, 51.06) mm, rotated rx 125.61 ry 0 rz 180 deg; joints [-9.737, -79.467, 124.305, 166.321, 45.662, -134.737]
  MoveL 280 to (0, -38.45, 51.06) mm, rotated rx 125.61 ry 0 rz 180 deg; joints [-8.34, -67.779, 108.621, 167.366, 41.538, -134.865]
  MoveL 281 to (0, -38.09, 51.53) mm, rotated rx 128.92 ry 0 rz 180 deg; joints [-8.968, -67.119, 108.853, 166.663, 42.513, -131.172]
  MoveL 282 to (-200, -38.09, 51.53) mm, rotated rx 128.92 ry 0 rz 180 deg; joints [-10.467, -78.668, 124.569, 165.574, 46.817, -131.1]
  MoveL 283 to (-200, -37.7, 51.99) mm, rotated rx 132.22 ry 0 rz 180 deg; joints [-11.151, -77.814, 124.836, 164.921, 48.022, -127.564]
  MoveL 284 to (0, -37.7, 51.99) mm, rotated rx 132.22 ry 0 rz 180 deg; joints [-9.558, -66.414, 109.088, 166.05, 43.53, -127.57]
  MoveL 285 to (0, -37.29, 52.42) mm, rotated rx 135.53 ry 0 rz 180 deg; joints [-10.108, -65.665, 109.325, 165.521, 44.585, -124.052]
  MoveL 286 to (-200, -37.29, 52.42) mm, rotated rx 135.53 ry 0 rz 180 deg; joints [-11.788, -76.906, 125.106, 164.36, 49.272, -124.121]
  MoveL 287 to (-200, -36.85, 52.83) mm, rotated rx 138.83 ry 0 rz 180 deg; joints [-12.378, -75.947, 125.377, 163.886, 50.56, -120.768]
  MoveL 288 to (0, -36.85, 52.83) mm, rotated rx 138.83 ry 0 rz 180 deg; joints [-10.618, -64.874, 109.563, 165.074, 45.672, -120.617]
  MoveL 289 to (0, -36.38, 53.21) mm, rotated rx 142.14 ry 0 rz 180 deg; joints [-11.084, -64.044, 109.799, 164.705, 46.786, -117.256]
  MoveL 290 to (-200, -36.38, 53.21) mm, rotated rx 142.14 ry 0 rz 180 deg; joints [-12.917, -74.939, 125.646, 163.493, 51.883, -117.496]
  MoveL 291 to (-200, -35.9, 53.56) mm, rotated rx 145.44 ry 0 rz 180 deg; joints [-13.405, -73.885, 125.911, 163.178, 53.234, -114.3]
  MoveL 292 to (0, -35.9, 53.56) mm, rotated rx 145.44 ry 0 rz 180 deg; joints [-11.507, -63.178, 110.031, 164.409, 47.924, -113.966]
  MoveL 293 to (0, -35.4, 53.89) mm, rotated rx 148.75 ry 0 rz 180 deg; joints [-11.885, -62.276, 110.26, 164.184, 49.081, -110.74]
  MoveL 294 to (-200, -35.4, 53.89) mm, rotated rx 148.75 ry 0 rz 180 deg; joints [-13.841, -72.787, 126.171, 162.936, 54.61, -111.171]
  MoveL 295 to (-200, -34.87, 54.19) mm, rotated rx 152.05 ry 0 rz 180 deg; joints [-14.224, -71.649, 126.424, 162.761, 56.006, -108.104]
  MoveL 296 to (0, -34.87, 54.19) mm, rotated rx 152.05 ry 0 rz 180 deg; joints [-12.218, -61.342, 110.483, 164.024, 50.254, -107.573]
  MoveL 297 to (0, -34.34, 54.45) mm, rotated rx 155.36 ry 0 rz 180 deg; joints [-12.503, -60.379, 110.699, 163.926, 51.438, -104.458]
  MoveL 298 to (-200, -34.34, 54.45) mm, rotated rx 155.36 ry 0 rz 180 deg; joints [-14.553, -70.474, 126.669, 162.65, 57.418, -105.09]
  MoveL 299 to (-200, -33.78, 54.69) mm, rotated rx 158.66 ry 0 rz 180 deg; joints [-14.827, -69.264, 126.904, 162.6, 58.841, -102.125]
  MoveL 300 to (0, -33.78, 54.69) mm, rotated rx 158.66 ry 0 rz 180 deg; joints [-12.742, -59.39, 110.906, 163.888, 52.63, -101.39]
  MoveL 301 to (0, -33.22, 54.89) mm, rotated rx 161.97 ry 0 rz 180 deg; joints [-12.932, -58.376, 111.104, 163.904, 53.826, -98.363]
  MoveL 302 to (-200, -33.22, 54.89) mm, rotated rx 161.97 ry 0 rz 180 deg; joints [-15.046, -68.025, 127.128, 162.606, 60.271, -99.199]
  MoveL 303 to (-200, -32.64, 55.06) mm, rotated rx 165.28 ry 0 rz 180 deg; joints [-15.21, -66.759, 127.339, 162.665, 61.706, -96.308]
  MoveL 304 to (0, -32.64, 55.06) mm, rotated rx 165.28 ry 0 rz 180 deg; joints [-13.075, -57.343, 111.292, 163.973, 55.023, -95.373]
  MoveL 305 to (0, -32.06, 55.19) mm, rotated rx 168.58 ry 0 rz 180 deg; joints [-13.169, -56.292, 111.468, 164.091, 56.218, -92.413]
  MoveL 306 to (-200, -32.06, 55.19) mm, rotated rx 168.58 ry 0 rz 180 deg; joints [-15.318, -65.47, 127.536, 162.775, 63.14, -93.444]
  MoveL 307 to (-200, -31.47, 55.3) mm, rotated rx 171.89 ry 0 rz 180 deg; joints [-15.37, -64.163, 127.719, 162.933, 64.571, -90.603]
  MoveL 308 to (0, -31.47, 55.3) mm, rotated rx 171.89 ry 0 rz 180 deg; joints [-13.214, -55.227, 111.632, 164.257, 57.407, -89.479]
  MoveL 309 to (0, -30.87, 55.36) mm, rotated rx 175.19 ry 0 rz 180 deg; joints [-13.211, -54.152, 111.784, 164.468, 58.588, -86.565]
  MoveL 310 to (-200, -30.87, 55.36) mm, rotated rx 175.19 ry 0 rz 180 deg; joints [-15.366, -62.842, 127.887, 163.138, 65.994, -87.777]
  MoveL 311 to (-200, -30.27, 55.4) mm, rotated rx 178.5 ry 0 rz 180 deg; joints [-15.306, -61.512, 128.038, 163.386, 67.406, -84.963]
  MoveL 312 to (0, -30.27, 55.4) mm, rotated rx 178.5 ry 0 rz 180 deg; joints [-13.159, -53.071, 111.922, 164.721, 59.756, -83.668]
  MoveL 313 to (0, -29.67, 55.4) mm, rotated rx 180 ry 0 rz 180 deg; joints [-13.119, -52.561, 111.981, 164.853, 60.301, -82.361]
  MoveL 314 to (-200, -29.67, 55.4) mm, rotated rx 180 ry 0 rz 180 deg; joints [-15.26, -60.884, 128.103, 163.516, 68.065, -83.692]
  MoveL 315 to (-200, -29.07, 55.4) mm, rotated rx 180 ry 0 rz 180 deg; joints [-15.26, -60.845, 128.105, 163.521, 68.104, -83.705]
  MoveL 316 to (0, -29.07, 55.4) mm, rotated rx 180 ry 0 rz 180 deg; joints [-13.119, -52.529, 111.984, 164.858, 60.333, -82.371]
  MoveL 317 to (0, -28.47, 55.4) mm, rotated rx 180 ry 0 rz 180 deg; joints [-13.119, -52.498, 111.986, 164.863, 60.365, -82.381]
  MoveL 318 to (-200, -28.47, 55.4) mm, rotated rx 180 ry 0 rz 180 deg; joints [-15.26, -60.807, 128.108, 163.526, 68.143, -83.717]
  MoveL 319 to (-200, -27.87, 55.4) mm, rotated rx 180 ry 0 rz 180 deg; joints [-15.26, -60.768, 128.11, 163.53, 68.182, -83.73]
  MoveL 320 to (0, -27.87, 55.4) mm, rotated rx 180 ry 0 rz 180 deg; joints [-13.119, -52.466, 111.988, 164.868, 60.397, -82.391]
  MoveL 321 to (0, -27.27, 55.4) mm, rotated rx 180 ry 0 rz 180 deg; joints [-13.119, -52.435, 111.99, 164.873, 60.43, -82.401]
  MoveL 322 to (-200, -27.27, 55.4) mm, rotated rx 180 ry 0 rz 180 deg; joints [-15.26, -60.73, 128.112, 163.535, 68.222, -83.742]
  MoveL 323 to (-200, -26.67, 55.4) mm, rotated rx 180 ry 0 rz 180 deg; joints [-15.26, -60.691, 128.114, 163.539, 68.261, -83.755]
  MoveL 324 to (0, -26.67, 55.4) mm, rotated rx 180 ry 0 rz 180 deg; joints [-13.119, -52.403, 111.992, 164.878, 60.462, -82.411]
  MoveL 325 to (0, -26.07, 55.4) mm, rotated rx 180 ry 0 rz 180 deg; joints [-13.119, -52.372, 111.994, 164.883, 60.494, -82.421]
  MoveL 326 to (-200, -26.07, 55.4) mm, rotated rx 180 ry 0 rz 180 deg; joints [-15.26, -60.652, 128.117, 163.544, 68.3, -83.767]
  MoveL 327 to (-200, -25.47, 55.4) mm, rotated rx 180 ry 0 rz 180 deg; joints [-15.26, -60.614, 128.119, 163.549, 68.339, -83.78]
  MoveL 328 to (0, -25.47, 55.4) mm, rotated rx 180 ry 0 rz 180 deg; joints [-13.119, -52.34, 111.996, 164.888, 60.527, -82.432]
  MoveL 329 to (0, -24.87, 55.4) mm, rotated rx 180 ry 0 rz 180 deg; joints [-13.119, -52.309, 111.997, 164.893, 60.559, -82.442]
  MoveL 330 to (-200, -24.87, 55.4) mm, rotated rx 180 ry 0 rz 180 deg; joints [-15.26, -60.575, 128.121, 163.553, 68.378, -83.792]
  MoveL 331 to (-200, -24.27, 55.4) mm, rotated rx 180 ry 0 rz 180 deg; joints [-15.26, -60.536, 128.123, 163.558, 68.417, -83.804]
  MoveL 332 to (0, -24.27, 55.4) mm, rotated rx 180 ry 0 rz 180 deg; joints [-13.119, -52.277, 111.999, 164.898, 60.591, -82.451]
  MoveL 333 to (0, -23.67, 55.4) mm, rotated rx 180 ry 0 rz 180 deg; joints [-13.119, -52.246, 112.001, 164.903, 60.623, -82.461]
  MoveL 334 to (-200, -23.67, 55.4) mm, rotated rx 180 ry 0 rz 180 deg; joints [-15.26, -60.498, 128.125, 163.562, 68.456, -83.817]
  MoveL 335 to (-200, -23.07, 55.4) mm, rotated rx 180 ry 0 rz 180 deg; joints [-15.26, -60.459, 128.127, 163.567, 68.495, -83.829]
  MoveL 336 to (0, -23.07, 55.4) mm, rotated rx 180 ry 0 rz 180 deg; joints [-13.119, -52.214, 112.003, 164.907, 60.656, -82.471]
  MoveL 337 to (0, -22.47, 55.4) mm, rotated rx 180 ry 0 rz 180 deg; joints [-13.119, -52.183, 112.005, 164.912, 60.688, -82.481]
  MoveL 338 to (-200, -22.47, 55.4) mm, rotated rx 180 ry 0 rz 180 deg; joints [-15.26, -60.42, 128.129, 163.571, 68.534, -83.842]
  MoveL 339 to (-200, -21.87, 55.4) mm, rotated rx 180 ry 0 rz 180 deg; joints [-15.26, -60.382, 128.131, 163.576, 68.573, -83.854]
  MoveL 340 to (0, -21.87, 55.4) mm, rotated rx 180 ry 0 rz 180 deg; joints [-13.119, -52.151, 112.007, 164.917, 60.72, -82.491]
  MoveL 341 to (0, -21.27, 55.4) mm, rotated rx 180 ry 0 rz 180 deg; joints [-13.119, -52.12, 112.008, 164.922, 60.752, -82.501]
  MoveL 342 to (-200, -21.27, 55.4) mm, rotated rx 180 ry 0 rz 180 deg; joints [-15.26, -60.343, 128.133, 163.58, 68.612, -83.866]
  MoveL 343 to (-200, -20.67, 55.4) mm, rotated rx 180 ry 0 rz 180 deg; joints [-15.26, -60.304, 128.135, 163.585, 68.651, -83.879]
  MoveL 344 to (0, -20.67, 55.4) mm, rotated rx 180 ry 0 rz 180 deg; joints [-13.119, -52.088, 112.01, 164.927, 60.784, -82.511]
  MoveL 345 to (0, -20.07, 55.4) mm, rotated rx 180 ry 0 rz 180 deg; joints [-13.119, -52.056, 112.012, 164.932, 60.816, -82.521]
  MoveL 346 to (-200, -20.07, 55.4) mm, rotated rx 180 ry 0 rz 180 deg; joints [-15.26, -60.265, 128.136, 163.589, 68.69, -83.891]
  MoveL 347 to (-200, -19.47, 55.4) mm, rotated rx 180 ry 0 rz 180 deg; joints [-15.26, -60.226, 128.138, 163.594, 68.729, -83.903]
  MoveL 348 to (0, -19.47, 55.4) mm, rotated rx 180 ry 0 rz 180 deg; joints [-13.119, -52.025, 112.013, 164.937, 60.848, -82.531]
  MoveL 349 to (0, -18.87, 55.4) mm, rotated rx 180 ry 0 rz 180 deg; joints [-13.119, -51.993, 112.015, 164.941, 60.881, -82.541]
  MoveL 350 to (-200, -18.87, 55.4) mm, rotated rx 180 ry 0 rz 180 deg; joints [-15.26, -60.187, 128.14, 163.598, 68.768, -83.916]
  MoveL 351 to (-200, -18.27, 55.4) mm, rotated rx 180 ry 0 rz 180 deg; joints [-15.26, -60.149, 128.142, 163.603, 68.807, -83.928]
  MoveL 352 to (0, -18.27, 55.4) mm, rotated rx 180 ry 0 rz 180 deg; joints [-13.119, -51.961, 112.016, 164.946, 60.913, -82.551]
  MoveL 353 to (0, -17.67, 55.4) mm, rotated rx 180 ry 0 rz 180 deg; joints [-13.119, -51.93, 112.018, 164.951, 60.945, -82.561]
  MoveL 354 to (-200, -17.67, 55.4) mm, rotated rx 180 ry 0 rz 180 deg; joints [-15.26, -60.11, 128.143, 163.607, 68.846, -83.94]
  MoveL 355 to (-200, -17.07, 55.4) mm, rotated rx 180 ry 0 rz 180 deg; joints [-15.26, -60.071, 128.145, 163.612, 68.885, -83.952]
  MoveL 356 to (0, -17.07, 55.4) mm, rotated rx 180 ry 0 rz 180 deg; joints [-13.119, -51.898, 112.019, 164.956, 60.977, -82.571]
  MoveL 357 to (0, -16.47, 55.4) mm, rotated rx 180 ry 0 rz 180 deg; joints [-13.119, -51.866, 112.021, 164.961, 61.009, -82.58]
  MoveL 358 to (-200, -16.47, 55.4) mm, rotated rx 180 ry 0 rz 180 deg; joints [-15.26, -60.032, 128.147, 163.616, 68.924, -83.965]
  MoveL 359 to (-200, -15.87, 55.4) mm, rotated rx 180 ry 0 rz 180 deg; joints [-15.26, -59.993, 128.148, 163.62, 68.963, -83.977]
  MoveL 360 to (0, -15.87, 55.4) mm, rotated rx 180 ry 0 rz 180 deg; joints [-13.119, -51.835, 112.022, 164.965, 61.041, -82.59]
  MoveL 361 to (0, -15.27, 55.4) mm, rotated rx 180 ry 0 rz 180 deg; joints [-13.119, -51.803, 112.024, 164.97, 61.073, -82.6]
  MoveL 362 to (-200, -15.27, 55.4) mm, rotated rx 180 ry 0 rz 180 deg; joints [-15.26, -59.954, 128.15, 163.625, 69.002, -83.989]
  MoveL 363 to (-200, -14.67, 55.4) mm, rotated rx 180 ry 0 rz 180 deg; joints [-15.26, -59.915, 128.151, 163.629, 69.041, -84.001]
  MoveL 364 to (0, -14.67, 55.4) mm, rotated rx 180 ry 0 rz 180 deg; joints [-13.119, -51.771, 112.025, 164.975, 61.105, -82.61]
  MoveL 365 to (0, -14.07, 55.4) mm, rotated rx 180 ry 0 rz 180 deg; joints [-13.119, -51.739, 112.027, 164.98, 61.137, -82.62]
  MoveL 366 to (-200, -14.07, 55.4) mm, rotated rx 180 ry 0 rz 180 deg; joints [-15.26, -59.876, 128.153, 163.634, 69.08, -84.014]
  MoveL 367 to (-200, -13.47, 55.4) mm, rotated rx 180 ry 0 rz 180 deg; joints [-15.26, -59.837, 128.154, 163.638, 69.118, -84.026]
  MoveL 368 to (0, -13.47, 55.4) mm, rotated rx 180 ry 0 rz 180 deg; joints [-13.119, -51.707, 112.028, 164.984, 61.169, -82.63]
  MoveL 369 to (0, -12.87, 55.4) mm, rotated rx 180 ry 0 rz 180 deg; joints [-13.119, -51.676, 112.029, 164.989, 61.201, -82.639]
  MoveL 370 to (-200, -12.87, 55.4) mm, rotated rx 180 ry 0 rz 180 deg; joints [-15.26, -59.798, 128.156, 163.642, 69.157, -84.038]
  MoveL 371 to (-200, -12.27, 55.4) mm, rotated rx 180 ry 0 rz 180 deg; joints [-15.26, -59.759, 128.157, 163.647, 69.196, -84.05]
  MoveL 372 to (0, -12.27, 55.4) mm, rotated rx 180 ry 0 rz 180 deg; joints [-13.119, -51.644, 112.03, 164.994, 61.233, -82.649]
  MoveL 373 to (0, -11.67, 55.4) mm, rotated rx 180 ry 0 rz 180 deg; joints [-13.119, -51.612, 112.032, 164.998, 61.265, -82.659]
  MoveL 374 to (-200, -11.67, 55.4) mm, rotated rx 180 ry 0 rz 180 deg; joints [-15.26, -59.72, 128.159, 163.651, 69.235, -84.062]
  MoveL 375 to (-200, -11.07, 55.4) mm, rotated rx 180 ry 0 rz 180 deg; joints [-15.26, -59.681, 128.16, 163.655, 69.274, -84.075]
  MoveL 376 to (0, -11.07, 55.4) mm, rotated rx 180 ry 0 rz 180 deg; joints [-13.119, -51.58, 112.033, 165.003, 61.297, -82.669]
  MoveL 377 to (0, -10.47, 55.4) mm, rotated rx 180 ry 0 rz 180 deg; joints [-13.119, -51.548, 112.034, 165.008, 61.329, -82.678]
  MoveL 378 to (-200, -10.47, 55.4) mm, rotated rx 180 ry 0 rz 180 deg; joints [-15.26, -59.642, 128.161, 163.66, 69.312, -84.087]
  MoveL 379 to (-200, -9.87, 55.4) mm, rotated rx 180 ry 0 rz 180 deg; joints [-15.26, -59.603, 128.163, 163.664, 69.351, -84.099]
  MoveL 380 to (0, -9.87, 55.4) mm, rotated rx 180 ry 0 rz 180 deg; joints [-13.119, -51.516, 112.035, 165.012, 61.361, -82.688]
  MoveL 381 to (0, -9.27, 55.4) mm, rotated rx 180 ry 0 rz 180 deg; joints [-13.119, -51.484, 112.036, 165.017, 61.393, -82.698]
  MoveL 382 to (-200, -9.27, 55.4) mm, rotated rx 180 ry 0 rz 180 deg; joints [-15.26, -59.564, 128.164, 163.668, 69.39, -84.111]
  MoveL 383 to (-200, -8.67, 55.4) mm, rotated rx 180 ry 0 rz 180 deg; joints [-15.26, -59.524, 128.165, 163.672, 69.429, -84.123]
  MoveL 384 to (0, -8.67, 55.4) mm, rotated rx 180 ry 0 rz 180 deg; joints [-13.119, -51.452, 112.037, 165.022, 61.425, -82.708]
  MoveL 385 to (0, -8.07, 55.4) mm, rotated rx 180 ry 0 rz 180 deg; joints [-13.119, -51.421, 112.038, 165.026, 61.457, -82.717]
  MoveL 386 to (-200, -8.07, 55.4) mm, rotated rx 180 ry 0 rz 180 deg; joints [-15.26, -59.485, 128.166, 163.677, 69.467, -84.135]
  MoveL 387 to (-200, -7.47, 55.4) mm, rotated rx 180 ry 0 rz 180 deg; joints [-15.26, -59.446, 128.167, 163.681, 69.506, -84.147]
  MoveL 388 to (0, -7.47, 55.4) mm, rotated rx 180 ry 0 rz 180 deg; joints [-13.119, -51.389, 112.04, 165.031, 61.488, -82.727]
  MoveL 389 to (0, -6.87, 55.4) mm, rotated rx 180 ry 0 rz 180 deg; joints [-13.119, -51.357, 112.041, 165.036, 61.52, -82.737]
  MoveL 390 to (-200, -6.87, 55.4) mm, rotated rx 180 ry 0 rz 180 deg; joints [-15.26, -59.407, 128.169, 163.685, 69.545, -84.159]
  MoveL 391 to (-200, -6.27, 55.4) mm, rotated rx 180 ry 0 rz 180 deg; joints [-15.26, -59.368, 128.17, 163.689, 69.583, -84.171]
  MoveL 392 to (0, -6.27, 55.4) mm, rotated rx 180 ry 0 rz 180 deg; joints [-13.119, -51.325, 112.042, 165.04, 61.552, -82.746]
  MoveL 393 to (0, -5.67, 55.4) mm, rotated rx 180 ry 0 rz 180 deg; joints [-13.119, -51.293, 112.042, 165.045, 61.584, -82.756]
  MoveL 394 to (-200, -5.67, 55.4) mm, rotated rx 180 ry 0 rz 180 deg; joints [-15.26, -59.328, 128.171, 163.694, 69.622, -84.184]
  MoveL 395 to (-200, -5.07, 55.4) mm, rotated rx 180 ry 0 rz 180 deg; joints [-15.26, -59.289, 128.172, 163.698, 69.661, -84.196]
  MoveL 396 to (0, -5.07, 55.4) mm, rotated rx 180 ry 0 rz 180 deg; joints [-13.119, -51.261, 112.043, 165.05, 61.616, -82.766]
  MoveL 397 to (0, -4.47, 55.4) mm, rotated rx 180 ry 0 rz 180 deg; joints [-13.119, -51.229, 112.044, 165.054, 61.648, -82.775]
  MoveL 398 to (-200, -4.47, 55.4) mm, rotated rx 180 ry 0 rz 180 deg; joints [-15.26, -59.25, 128.173, 163.702, 69.699, -84.208]
  MoveL 399 to (-200, -3.87, 55.4) mm, rotated rx 180 ry 0 rz 180 deg; joints [-15.26, -59.211, 128.174, 163.706, 69.738, -84.22]
  MoveL 400 to (0, -3.87, 55.4) mm, rotated rx 180 ry 0 rz 180 deg; joints [-13.119, -51.197, 112.045, 165.059, 61.679, -82.785]
  MoveL 401 to (0, -3.27, 55.4) mm, rotated rx 180 ry 0 rz 180 deg; joints [-13.119, -51.164, 112.046, 165.063, 61.711, -82.795]
  MoveL 402 to (-200, -3.27, 55.4) mm, rotated rx 180 ry 0 rz 180 deg; joints [-15.26, -59.171, 128.175, 163.71, 69.777, -84.232]
  MoveL 403 to (-200, -2.67, 55.4) mm, rotated rx 180 ry 0 rz 180 deg; joints [-15.26, -59.132, 128.175, 163.714, 69.815, -84.244]
  MoveL 404 to (0, -2.67, 55.4) mm, rotated rx 180 ry 0 rz 180 deg; joints [-13.119, -51.132, 112.047, 165.068, 61.743, -82.804]
  MoveL 405 to (0, -2.07, 55.4) mm, rotated rx 180 ry 0 rz 180 deg; joints [-13.119, -51.1, 112.047, 165.072, 61.775, -82.814]
  MoveL 406 to (-200, -2.07, 55.4) mm, rotated rx 180 ry 0 rz 180 deg; joints [-15.26, -59.093, 128.176, 163.719, 69.854, -84.256]
  MoveL 407 to (-200, -1.47, 55.4) mm, rotated rx 180 ry 0 rz 180 deg; joints [-15.26, -59.053, 128.177, 163.723, 69.892, -84.268]
  MoveL 408 to (0, -1.47, 55.4) mm, rotated rx 180 ry 0 rz 180 deg; joints [-13.119, -51.068, 112.048, 165.077, 61.806, -82.823]
  MoveL 409 to (0, -0.87, 55.4) mm, rotated rx 180 ry 0 rz 180 deg; joints [-13.119, -51.036, 112.049, 165.081, 61.838, -82.833]
  MoveL 410 to (-200, -0.87, 55.4) mm, rotated rx 180 ry 0 rz 180 deg; joints [-15.26, -59.014, 128.178, 163.727, 69.931, -84.28]
  MoveL 411 to (-200, -0.27, 55.4) mm, rotated rx 180 ry 0 rz 180 deg; joints [-15.26, -58.975, 128.179, 163.731, 69.969, -84.292]
  MoveL 412 to (0, -0.27, 55.4) mm, rotated rx 180 ry 0 rz 180 deg; joints [-13.119, -51.004, 112.05, 165.086, 61.87, -82.843]
  MoveL 413 to (0, 0, 55.4) mm, rotated rx 180 ry 0 rz 180 deg; joints [-13.119, -50.989, 112.05, 165.088, 61.884, -82.847]
  MoveL 414 to (-200, 0, 55.4) mm, rotated rx 180 ry 0 rz 180 deg; joints [-15.26, -58.957, 128.179, 163.733, 69.987, -84.297]
  MoveL 415 to (-200, 0, 55.8) mm, rotated rx 180 ry 0 rz 180 deg; joints [-15.278, -58.953, 128.171, 163.713, 69.985, -84.289]
  MoveL 416 to (0, 0, 55.8) mm, rotated rx 180 ry 0 rz 180 deg; joints [-13.135, -50.985, 112.042, 165.07, 61.882, -82.837]
  MoveL 417 to (0, -0.6, 55.8) mm, rotated rx 180 ry 0 rz 180 deg; joints [-13.135, -51.017, 112.041, 165.065, 61.851, -82.828]
  MoveL 418 to (-200, -0.6, 55.8) mm, rotated rx 180 ry 0 rz 180 deg; joints [-15.278, -58.992, 128.17, 163.709, 69.946, -84.277]
  MoveL 419 to (-200, -1.2, 55.8) mm, rotated rx 180 ry 0 rz 180 deg; joints [-15.278, -59.031, 128.169, 163.705, 69.908, -84.265]
  MoveL 420 to (0, -1.2, 55.8) mm, rotated rx 180 ry 0 rz 180 deg; joints [-13.135, -51.05, 112.041, 165.061, 61.819, -82.818]
  MoveL 421 to (0, -1.8, 55.8) mm, rotated rx 180 ry 0 rz 180 deg; joints [-13.135, -51.082, 112.04, 165.056, 61.787, -82.809]
  MoveL 422 to (-200, -1.8, 55.8) mm, rotated rx 180 ry 0 rz 180 deg; joints [-15.278, -59.071, 128.168, 163.701, 69.869, -84.253]
  MoveL 423 to (-200, -2.4, 55.8) mm, rotated rx 180 ry 0 rz 180 deg; joints [-15.278, -59.11, 128.167, 163.697, 69.83, -84.241]
  MoveL 424 to (0, -2.4, 55.8) mm, rotated rx 180 ry 0 rz 180 deg; joints [-13.135, -51.114, 112.039, 165.051, 61.755, -82.799]
  MoveL 425 to (0, -3, 55.8) mm, rotated rx 180 ry 0 rz 180 deg; joints [-13.135, -51.146, 112.038, 165.047, 61.724, -82.789]
  MoveL 426 to (-200, -3, 55.8) mm, rotated rx 180 ry 0 rz 180 deg; joints [-15.278, -59.149, 128.167, 163.692, 69.792, -84.229]
  MoveL 427 to (-200, -3.6, 55.8) mm, rotated rx 180 ry 0 rz 180 deg; joints [-15.278, -59.189, 128.166, 163.688, 69.753, -84.217]
  MoveL 428 to (0, -3.6, 55.8) mm, rotated rx 180 ry 0 rz 180 deg; joints [-13.135, -51.178, 112.038, 165.042, 61.692, -82.78]
  MoveL 429 to (0, -4.2, 55.8) mm, rotated rx 180 ry 0 rz 180 deg; joints [-13.135, -51.21, 112.037, 165.038, 61.66, -82.77]
  MoveL 430 to (-200, -4.2, 55.8) mm, rotated rx 180 ry 0 rz 180 deg; joints [-15.278, -59.228, 128.165, 163.684, 69.715, -84.205]
  MoveL 431 to (-200, -4.8, 55.8) mm, rotated rx 180 ry 0 rz 180 deg; joints [-15.278, -59.267, 128.164, 163.68, 69.676, -84.193]
  MoveL 432 to (0, -4.8, 55.8) mm, rotated rx 180 ry 0 rz 180 deg; joints [-13.135, -51.242, 112.036, 165.033, 61.628, -82.76]
  MoveL 433 to (0, -5.4, 55.8) mm, rotated rx 180 ry 0 rz 180 deg; joints [-13.135, -51.274, 112.035, 165.029, 61.597, -82.751]
  MoveL 434 to (-200, -5.4, 55.8) mm, rotated rx 180 ry 0 rz 180 deg; joints [-15.278, -59.306, 128.163, 163.676, 69.637, -84.181]
  MoveL 435 to (-200, -6, 55.8) mm, rotated rx 180 ry 0 rz 180 deg; joints [-15.278, -59.346, 128.162, 163.671, 69.599, -84.169]
  MoveL 436 to (0, -6, 55.8) mm, rotated rx 180 ry 0 rz 180 deg; joints [-13.135, -51.306, 112.034, 165.024, 61.565, -82.741]
  MoveL 437 to (0, -6.6, 55.8) mm, rotated rx 180 ry 0 rz 180 deg; joints [-13.135, -51.338, 112.033, 165.019, 61.533, -82.731]
  MoveL 438 to (-200, -6.6, 55.8) mm, rotated rx 180 ry 0 rz 180 deg; joints [-15.278, -59.385, 128.161, 163.667, 69.56, -84.157]
  MoveL 439 to (-200, -7.2, 55.8) mm, rotated rx 180 ry 0 rz 180 deg; joints [-15.278, -59.424, 128.16, 163.663, 69.521, -84.145]
  MoveL 440 to (0, -7.2, 55.8) mm, rotated rx 180 ry 0 rz 180 deg; joints [-13.135, -51.37, 112.032, 165.015, 61.501, -82.722]
  MoveL 441 to (0, -7.8, 55.8) mm, rotated rx 180 ry 0 rz 180 deg; joints [-13.135, -51.402, 112.031, 165.01, 61.469, -82.712]
  MoveL 442 to (-200, -7.8, 55.8) mm, rotated rx 180 ry 0 rz 180 deg; joints [-15.278, -59.463, 128.158, 163.659, 69.483, -84.133]
  MoveL 443 to (-200, -8.4, 55.8) mm, rotated rx 180 ry 0 rz 180 deg; joints [-15.278, -59.502, 128.157, 163.655, 69.444, -84.121]
  MoveL 444 to (0, -8.4, 55.8) mm, rotated rx 180 ry 0 rz 180 deg; joints [-13.135, -51.434, 112.03, 165.005, 61.437, -82.702]
  MoveL 445 to (0, -9, 55.8) mm, rotated rx 180 ry 0 rz 180 deg; joints [-13.135, -51.466, 112.029, 165.001, 61.405, -82.693]
  MoveL 446 to (-200, -9, 55.8) mm, rotated rx 180 ry 0 rz 180 deg; joints [-15.278, -59.542, 128.156, 163.65, 69.405, -84.108]
  MoveL 447 to (-200, -9.6, 55.8) mm, rotated rx 180 ry 0 rz 180 deg; joints [-15.278, -59.581, 128.155, 163.646, 69.367, -84.096]
  MoveL 448 to (0, -9.6, 55.8) mm, rotated rx 180 ry 0 rz 180 deg; joints [-13.135, -51.498, 112.028, 164.996, 61.374, -82.683]
  MoveL 449 to (0, -10.2, 55.8) mm, rotated rx 180 ry 0 rz 180 deg; joints [-13.135, -51.53, 112.027, 164.991, 61.342, -82.673]
  MoveL 450 to (-200, -10.2, 55.8) mm, rotated rx 180 ry 0 rz 180 deg; joints [-15.278, -59.62, 128.154, 163.642, 69.328, -84.084]
  MoveL 451 to (-200, -10.8, 55.8) mm, rotated rx 180 ry 0 rz 180 deg; joints [-15.278, -59.659, 128.152, 163.637, 69.289, -84.072]
  MoveL 452 to (0, -10.8, 55.8) mm, rotated rx 180 ry 0 rz 180 deg; joints [-13.135, -51.562, 112.025, 164.987, 61.31, -82.663]
  MoveL 453 to (0, -11.4, 55.8) mm, rotated rx 180 ry 0 rz 180 deg; joints [-13.135, -51.593, 112.024, 164.982, 61.278, -82.654]
  MoveL 454 to (-200, -11.4, 55.8) mm, rotated rx 180 ry 0 rz 180 deg; joints [-15.278, -59.698, 128.151, 163.633, 69.25, -84.06]
  MoveL 455 to (-200, -12, 55.8) mm, rotated rx 180 ry 0 rz 180 deg; joints [-15.278, -59.737, 128.15, 163.629, 69.212, -84.048]
  MoveL 456 to (0, -12, 55.8) mm, rotated rx 180 ry 0 rz 180 deg; joints [-13.135, -51.625, 112.023, 164.977, 61.246, -82.644]
  MoveL 457 to (0, -12.6, 55.8) mm, rotated rx 180 ry 0 rz 180 deg; joints [-13.135, -51.657, 112.022, 164.973, 61.214, -82.634]
  MoveL 458 to (-200, -12.6, 55.8) mm, rotated rx 180 ry 0 rz 180 deg; joints [-15.278, -59.776, 128.148, 163.624, 69.173, -84.035]
  MoveL 459 to (-200, -13.2, 55.8) mm, rotated rx 180 ry 0 rz 180 deg; joints [-15.278, -59.815, 128.147, 163.62, 69.134, -84.023]
  MoveL 460 to (0, -13.2, 55.8) mm, rotated rx 180 ry 0 rz 180 deg; joints [-13.135, -51.689, 112.02, 164.968, 61.182, -82.624]
  MoveL 461 to (0, -13.8, 55.8) mm, rotated rx 180 ry 0 rz 180 deg; joints [-13.135, -51.721, 112.019, 164.963, 61.15, -82.614]
  MoveL 462 to (-200, -13.8, 55.8) mm, rotated rx 180 ry 0 rz 180 deg; joints [-15.278, -59.854, 128.145, 163.616, 69.095, -84.011]
  MoveL 463 to (-200, -14.4, 55.8) mm, rotated rx 180 ry 0 rz 180 deg; joints [-15.278, -59.893, 128.144, 163.611, 69.056, -83.999]
  MoveL 464 to (0, -14.4, 55.8) mm, rotated rx 180 ry 0 rz 180 deg; joints [-13.135, -51.753, 112.018, 164.959, 61.118, -82.605]
  MoveL 465 to (0, -15, 55.8) mm, rotated rx 180 ry 0 rz 180 deg; joints [-13.135, -51.784, 112.016, 164.954, 61.086, -82.595]
  MoveL 466 to (-200, -15, 55.8) mm, rotated rx 180 ry 0 rz 180 deg; joints [-15.278, -59.932, 128.142, 163.607, 69.017, -83.987]
  MoveL 467 to (-200, -15.6, 55.8) mm, rotated rx 180 ry 0 rz 180 deg; joints [-15.278, -59.971, 128.141, 163.603, 68.979, -83.974]
  MoveL 468 to (0, -15.6, 55.8) mm, rotated rx 180 ry 0 rz 180 deg; joints [-13.135, -51.816, 112.015, 164.949, 61.054, -82.585]
  MoveL 469 to (0, -16.2, 55.8) mm, rotated rx 180 ry 0 rz 180 deg; joints [-13.135, -51.848, 112.014, 164.944, 61.022, -82.575]
  MoveL 470 to (-200, -16.2, 55.8) mm, rotated rx 180 ry 0 rz 180 deg; joints [-15.278, -60.01, 128.139, 163.598, 68.94, -83.962]
  MoveL 471 to (-200, -16.8, 55.8) mm, rotated rx 180 ry 0 rz 180 deg; joints [-15.278, -60.049, 128.138, 163.594, 68.901, -83.95]
  MoveL 472 to (0, -16.8, 55.8) mm, rotated rx 180 ry 0 rz 180 deg; joints [-13.135, -51.88, 112.012, 164.939, 60.99, -82.565]
  MoveL 473 to (0, -17.4, 55.8) mm, rotated rx 180 ry 0 rz 180 deg; joints [-13.135, -51.911, 112.011, 164.935, 60.958, -82.555]
  MoveL 474 to (-200, -17.4, 55.8) mm, rotated rx 180 ry 0 rz 180 deg; joints [-15.278, -60.088, 128.136, 163.589, 68.862, -83.937]
  MoveL 475 to (-200, -18, 55.8) mm, rotated rx 180 ry 0 rz 180 deg; joints [-15.278, -60.127, 128.134, 163.585, 68.823, -83.925]
  MoveL 476 to (0, -18, 55.8) mm, rotated rx 180 ry 0 rz 180 deg; joints [-13.135, -51.943, 112.009, 164.93, 60.926, -82.545]
  MoveL 477 to (0, -18.6, 55.8) mm, rotated rx 180 ry 0 rz 180 deg; joints [-13.135, -51.975, 112.008, 164.925, 60.893, -82.536]
  MoveL 478 to (-200, -18.6, 55.8) mm, rotated rx 180 ry 0 rz 180 deg; joints [-15.278, -60.166, 128.132, 163.581, 68.784, -83.913]
  MoveL 479 to (-200, -19.2, 55.8) mm, rotated rx 180 ry 0 rz 180 deg; joints [-15.278, -60.204, 128.131, 163.576, 68.745, -83.901]
  MoveL 480 to (0, -19.2, 55.8) mm, rotated rx 180 ry 0 rz 180 deg; joints [-13.135, -52.006, 112.006, 164.92, 60.861, -82.526]
  MoveL 481 to (0, -19.8, 55.8) mm, rotated rx 180 ry 0 rz 180 deg; joints [-13.135, -52.038, 112.004, 164.915, 60.829, -82.516]
  MoveL 482 to (-200, -19.8, 55.8) mm, rotated rx 180 ry 0 rz 180 deg; joints [-15.278, -60.243, 128.129, 163.572, 68.706, -83.888]
  MoveL 483 to (-200, -20.4, 55.8) mm, rotated rx 180 ry 0 rz 180 deg; joints [-15.278, -60.282, 128.127, 163.567, 68.667, -83.876]
  MoveL 484 to (0, -20.4, 55.8) mm, rotated rx 180 ry 0 rz 180 deg; joints [-13.135, -52.07, 112.003, 164.911, 60.797, -82.506]
  MoveL 485 to (0, -21, 55.8) mm, rotated rx 180 ry 0 rz 180 deg; joints [-13.135, -52.101, 112.001, 164.906, 60.765, -82.496]
  MoveL 486 to (-200, -21, 55.8) mm, rotated rx 180 ry 0 rz 180 deg; joints [-15.278, -60.321, 128.125, 163.563, 68.628, -83.864]
  MoveL 487 to (-200, -21.6, 55.8) mm, rotated rx 180 ry 0 rz 180 deg; joints [-15.278, -60.36, 128.123, 163.558, 68.589, -83.851]
  MoveL 488 to (0, -21.6, 55.8) mm, rotated rx 180 ry 0 rz 180 deg; joints [-13.135, -52.133, 111.999, 164.901, 60.733, -82.486]
  MoveL 489 to (0, -22.2, 55.8) mm, rotated rx 180 ry 0 rz 180 deg; joints [-13.135, -52.164, 111.998, 164.896, 60.701, -82.476]
  MoveL 490 to (-200, -22.2, 55.8) mm, rotated rx 180 ry 0 rz 180 deg; joints [-15.278, -60.398, 128.121, 163.554, 68.55, -83.839]
  MoveL 491 to (-200, -22.8, 55.8) mm, rotated rx 180 ry 0 rz 180 deg; joints [-15.278, -60.437, 128.119, 163.549, 68.511, -83.826]
  MoveL 492 to (0, -22.8, 55.8) mm, rotated rx 180 ry 0 rz 180 deg; joints [-13.135, -52.196, 111.996, 164.891, 60.668, -82.466]
  MoveL 493 to (0, -23.4, 55.8) mm, rotated rx 180 ry 0 rz 180 deg; joints [-13.135, -52.228, 111.994, 164.886, 60.636, -82.456]
  MoveL 494 to (-200, -23.4, 55.8) mm, rotated rx 180 ry 0 rz 180 deg; joints [-15.278, -60.476, 128.117, 163.545, 68.472, -83.814]
  MoveL 495 to (-200, -24, 55.8) mm, rotated rx 180 ry 0 rz 180 deg; joints [-15.278, -60.515, 128.115, 163.54, 68.433, -83.802]
  MoveL 496 to (0, -24, 55.8) mm, rotated rx 180 ry 0 rz 180 deg; joints [-13.135, -52.259, 111.992, 164.881, 60.604, -82.446]
  MoveL 497 to (0, -24.6, 55.8) mm, rotated rx 180 ry 0 rz 180 deg; joints [-13.135, -52.291, 111.99, 164.876, 60.572, -82.436]
  MoveL 498 to (-200, -24.6, 55.8) mm, rotated rx 180 ry 0 rz 180 deg; joints [-15.278, -60.553, 128.113, 163.535, 68.394, -83.789]
  MoveL 499 to (-200, -25.2, 55.8) mm, rotated rx 180 ry 0 rz 180 deg; joints [-15.278, -60.592, 128.111, 163.531, 68.355, -83.777]
  MoveL 500 to (0, -25.2, 55.8) mm, rotated rx 180 ry 0 rz 180 deg; joints [-13.135, -52.322, 111.988, 164.871, 60.54, -82.426]
  MoveL 501 to (0, -25.8, 55.8) mm, rotated rx 180 ry 0 rz 180 deg; joints [-13.135, -52.354, 111.987, 164.867, 60.507, -82.416]
  MoveL 502 to (-200, -25.8, 55.8) mm, rotated rx 180 ry 0 rz 180 deg; joints [-15.278, -60.631, 128.109, 163.526, 68.316, -83.764]
  MoveL 503 to (-200, -26.4, 55.8) mm, rotated rx 180 ry 0 rz 180 deg; joints [-15.278, -60.669, 128.107, 163.522, 68.277, -83.752]
  MoveL 504 to (0, -26.4, 55.8) mm, rotated rx 180 ry 0 rz 180 deg; joints [-13.135, -52.385, 111.985, 164.862, 60.475, -82.406]
  MoveL 505 to (0, -27, 55.8) mm, rotated rx 180 ry 0 rz 180 deg; joints [-13.135, -52.417, 111.983, 164.857, 60.443, -82.396]
  MoveL 506 to (-200, -27, 55.8) mm, rotated rx 180 ry 0 rz 180 deg; joints [-15.278, -60.708, 128.105, 163.517, 68.238, -83.739]
  MoveL 507 to (-200, -27.6, 55.8) mm, rotated rx 180 ry 0 rz 180 deg; joints [-15.278, -60.746, 128.103, 163.512, 68.198, -83.727]
  MoveL 508 to (0, -27.6, 55.8) mm, rotated rx 180 ry 0 rz 180 deg; joints [-13.135, -52.448, 111.981, 164.852, 60.411, -82.386]
  MoveL 509 to (0, -28.2, 55.8) mm, rotated rx 180 ry 0 rz 180 deg; joints [-13.135, -52.479, 111.979, 164.847, 60.378, -82.376]
  MoveL 510 to (-200, -28.2, 55.8) mm, rotated rx 180 ry 0 rz 180 deg; joints [-15.278, -60.785, 128.1, 163.508, 68.159, -83.714]
  MoveL 511 to (-200, -28.8, 55.8) mm, rotated rx 180 ry 0 rz 180 deg; joints [-15.278, -60.824, 128.098, 163.503, 68.12, -83.702]
  MoveL 512 to (0, -28.8, 55.8) mm, rotated rx 180 ry 0 rz 180 deg; joints [-13.135, -52.511, 111.977, 164.842, 60.346, -82.366]
  MoveL 513 to (0, -29.4, 55.8) mm, rotated rx 180 ry 0 rz 180 deg; joints [-13.135, -52.542, 111.974, 164.837, 60.314, -82.356]
  MoveL 514 to (-200, -29.4, 55.8) mm, rotated rx 180 ry 0 rz 180 deg; joints [-15.278, -60.862, 128.096, 163.498, 68.081, -83.689]
  MoveL 515 to (-200, -30, 55.8) mm, rotated rx 180 ry 0 rz 180 deg; joints [-15.278, -60.901, 128.093, 163.494, 68.042, -83.677]
  MoveL 516 to (0, -30, 55.8) mm, rotated rx 180 ry 0 rz 180 deg; joints [-13.135, -52.574, 111.972, 164.832, 60.281, -82.346]
  MoveL 517 to (0, -30.6, 55.78) mm, rotated rx 176.82 ry 0 rz 180 deg; joints [-13.207, -53.618, 111.845, 164.568, 59.161, -85.129]
  MoveL 518 to (-200, -30.6, 55.78) mm, rotated rx 176.82 ry 0 rz 180 deg; joints [-15.362, -62.186, 127.955, 163.234, 66.687, -86.384]
  MoveL 519 to (-200, -31.2, 55.73) mm, rotated rx 173.63 ry 0 rz 180 deg; joints [-15.393, -63.465, 127.801, 163.015, 65.32, -89.098]
  MoveL 520 to (0, -31.2, 55.73) mm, rotated rx 173.63 ry 0 rz 180 deg; joints [-13.234, -54.658, 111.706, 164.344, 58.029, -87.925]
